text list "Input_注释": 0 '备用'; 1 '备用'; 2 '备用'; 3 '备用'; 4 '备用'; 5 '备用'; 6 '备用'; 7 '备用'; 10 '备用'; 11 '备用'; 12 '备用'; 13 '备用'; 14 '备用'; 15 '备用'; 16 '备用'; 17 '备用'; 20 '紧急停止 / 备用'; 21 '总气压检测 / 备用'; 22 '手动模式 / 备用'; 23 '自动模式 / 备用'; 24 '启动运行按钮 / 备用'; 25 '故障复位按钮 / 备用'; 26 '启动按钮输入 / 备用'; 27 '光幕Ok / RobotReadyToMark'; 30 '旁路钥匙开关'; 31 '备用 / RobotTrayFullToOut'; 32 '变频器Ready / RobotPartInTurner'; 33 '备用 / reserve'; 34 '备用'; 35 '备用'; 36 '备用'; 37 '备用'; 40 '备用'; 41 '备用'; 42 '备用'; 43 '备用'; 44 '备用'; 45 '备用'; 46 '备用'; 47 '备用'; 50 '备用'; 51 '备用'; 52 '备用'; 53 '备用'; 54 '备用'; 55 '备用'; 56 '备用'; 57 '备用'; 200 '10插销缸缩回位磁开 / Communication with Conveyor / 与Conveyor通讯'; 201 '10插销缸伸出位磁开 / Communication with Conveyor / 与Conveyor通讯'; 202 '10测试滑台缸伸出位磁开'; 203 '10测试滑台缸缩回位磁开 / Communication with Conveyor / 与Conveyor通讯'; 204 '10测试升降缸伸出位磁开 / Communication with Conveyor / 与Conveyor通讯'; 205 '10测试升降缸缩回位磁开 / Communication with Conveyor / 与Conveyor通讯'; 206 '10滑台推出缸缩回位磁开 / Communication with Conveyor / 与Conveyor通讯'; 207 '10滑台推出缸伸出位磁开 / Communication with Conveyor / 与Conveyor通讯'; 210 '10下料滑台缸伸出位磁开 / Communication with Conveyor / 与Conveyor通讯'; 211 '10下料滑台缸缩回位磁开 / Communication with Conveyor / 与Conveyor通讯'; 212 '11下料升降缸伸出位磁开 / Communication with Conveyor / 与Conveyor通讯'; 213 '11下料升降缸缩回位磁开 / Communication with Conveyor / 与Conveyor通讯'; 214 '11下料夹爪缸伸出位磁开 / Communication with Conveyor / 与Conveyor通讯'; 215 '11下料夹爪缸缩回位磁开 / Communication with Conveyor / 与Conveyor通讯'; 216 '11废料阻挡缸伸出位磁开 / Communication with Conveyor / 与Conveyor通讯'; 217 '11废料阻挡缸缩回位磁开 / Communication with Conveyor / 与Conveyor通讯'; 222 '10.气密工件到位接近开关信号 / Communication with Conveyor / 与Conveyor通讯'; 223 '10.废料检测信号 / Communication with Conveyor / 与Conveyor通讯'; 224 '11.气密下料工件到位信号 / Communication with Conveyor / 与Conveyor通讯'; 225 '备用 / Communication with Conveyor / 与Conveyor通讯'; 226 '备用 / Communication with Conveyor / 与Conveyor通讯'; 227 '备用 / Communication with Conveyor / 与Conveyor通讯'; 230 '2垂直探针缸伸出位磁开 / Communication with Conveyor / 与Conveyor通讯'; 232 '备用 / Communication with Conveyor / 与Conveyor通讯'; 233 '备用 / Communication with Conveyor / 与Conveyor通讯'; 234 '转盘上料位工件到位信号 / Communication with Conveyor / 与Conveyor通讯'; 235 '备用 / Communication with Conveyor / 与Conveyor通讯'; 236 '备用 / Communication with Conveyor / 与Conveyor通讯'; 240 '2水平探针缸伸出位磁开 / Indexing plate number 3 / 转盘编号3'; 241 '2水平探针缸缩回位磁开 / Indexing plate number 4 / 转盘编号4'; 242 '8升降缸伸出位磁开 / 06.压紧缸原点位磁开'; 243 '8升降缸缩回位磁开 / 06.压紧缸工作位磁开'; 244 '2夹紧缸缩回位磁开 / 06.热烫缸原点位磁开'; 245 '2夹紧缸伸出位磁开 / 06.热烫缸工作位磁开'; 246 '备用 / 02.升降缸原点位磁开'; 247 '备用 / 02.升降缸工作位磁开'; 250 '4齿面凹面转换缸伸出位磁开 / Indexing plate number 1 / 转盘编号1'; 251 '4齿面凹面转换缸缩回位磁开 / Indexing plate number 2 / 转盘编号2'; 252 '4垂直探针缸伸出位磁开 / 上料托盘检测光电1'; 253 '4垂直探针缸缩回位磁开 / 上料皮带挡料1缸工作位磁开'; 254 '4夹紧缸缩回位磁开 / 上料皮带挡料2缸工作位磁开'; 255 '4夹紧缸伸出位磁开 / 上料托盘检测光电2'; 256 '4水平探针缸伸出位磁开 / 02.送料长缸工作位磁开'; 257 '4水平探针缸缩回位磁开 / 02.送料长缸原点位磁开'; 260 '6夹紧缸缩回位磁开 / 02.送料短缸工作位磁开'; 261 '6夹紧缸伸出位磁开 / 01.真空*工作位磁开'; 262 '6水平探针缸伸出位磁开 / 06.热烫缸工作位磁开'; 263 '6水平探针缸缩回位磁开 / 06.热烫缸工作位磁开'; 264 '6垂直探针缸伸出位磁开 / 06.热烫缸工作位磁开'; 265 '6垂直探针缸缩回位磁开 / 06.热烫缸工作位磁开'; 266 '02.转台编码 Bit0 / 06.热烫缸工作位磁开'; 267 '02.转台编码 Bit1 / 06.热烫缸工作位磁开'; 270 '02.转台编码 Bit2 / 06.热烫缸工作位磁开'; 271 '02.转台编码 Bit3 / 06.热烫缸工作位磁开'; 272 '备用 / 06.热烫缸工作位磁开'; 273 '备用 / 06.热烫缸工作位磁开'; 274 '备用 / 06.热烫缸工作位磁开'; 275 '备用 / 06.热烫缸工作位磁开'; 276 '备用 / 06.热烫缸工作位磁开'; 277 '备用 / 06.热烫缸工作位磁开'; 280 '备用 / 06.热烫缸工作位磁开'; 220 '10.气密工件到位光电信号 / Communication with Conveyor / 与Conveyor通讯'; 221 '备用 / Communication with Conveyor / 与Conveyor通讯'; 231 '2垂直探针缸缩回位磁开 / Communication with Conveyor / 与Conveyor通讯'; 237 '转台到位检测接近 / Communication with Conveyor / 与Conveyor通讯'; 281 '备用 / 06.热烫缸工作位磁开'; 282 '备用 / 06.热烫缸工作位磁开'; 283 '备用 / 06.热烫缸工作位磁开'; 284 '备用 / 06.热烫缸工作位磁开'; 285 '备用 / 06.热烫缸工作位磁开'; 286 '07.工件到位信号'; 287 '备用'; 290 '07.插销缸缩回信号'; 291 '07.插销缸伸出信号'; 292 '07.压紧缸缩回信号'; 293 '07.压紧缸伸出信号'; 294 '备用'; 295 '备用'; 296 '07.滑台推进缸伸出信号'; 297 '07.滑台推进缸缩回信号'; 300 '07.下料滑台缸缩回信号'; 301 '07.下料滑台缸伸出信号'; 302 '08.下料升降缸伸出信号'; 303 '08.下料升降缸缩回信号'; 304 '08.下料夹爪缸缩回信号'; 305 '08.下料夹爪缸伸出信号'; 306 '08.下料止挡缸伸出信号'; 307 '08.下料止挡缸缩回信号'; 310 '备用'; 311 '备用'; 312 '备用'; 313 '备用'; 314 '备用'; 315 '备用'; 316 '备用'; 317 '备用'; 74 '备用'; 77 '备用'; 76 '备用'; 75 '备用'; 73 '备用'; 72 '备用'; 71 '备用'; 70 '备用'; 67 '备用'; 66 '备用'; 65 '备用'; 64 '备用'; 63 '备用'; 62 '备用'; 61 '备用'; 60 '备用'; 320 '备用'; 321 '备用'; 322 '备用'; 323 '备用'; 324 '备用'; 325 '备用'; 326 '备用'; 327 '备用'; 330 '备用'; 331 '备用'; 332 '备用'; 333 '备用'; 334 '备用'; 335 '备用'; 336 '备用'; 337 '备用'; 340 '备用'; 341 '备用'; 342 '备用'; 343 '备用'; 344 '备用'; 345 '备用'; 346 '备用'; 347 '备用'; 350 '备用'; 351 '备用'; 352 '备用'; 353 '备用'; 354 '备用'; 355 '备用'; 356 '备用'; 357 '备用'

text list "OutPut_地址": 0 'Q0.0'; 1 'Q0.1'; 2 'Q0.2'; 3 'Q0.3'; 4 'Q0.4'; 5 'Q0.5'; 6 'Q0.6'; 7 'Q0.7'; 10 'Q1.0'; 11 'Q1.1'; 12 'Q1.2'; 13 'Q1.3'; 14 'Q1.4'; 15 'Q1.5'; 16 'Q1.6'; 17 'Q1.7'; 20 'Q2.0'; 21 'Q2.1'; 22 'Q2.2'; 23 'Q2.3'; 24 'Q2.4'; 25 'Q2.5'; 26 'Q2.6'; 27 'Q2.7'; 30 'Q3.0'; 31 'Q3.1'; 32 'Q3.2'; 33 'Q3.3'; 34 'Q3.4'; 35 'Q3.5'; 36 'Q3.6'; 37 'Q3.7'; 40 'Q4.0'; 41 'Q4.1'; 42 'Q4.2'; 43 'Q4.3'; 44 'Q4.4'; 45 'Q4.5'; 46 'Q4.6'; 47 'Q4.7'; 50 'Q5.0'; 51 'Q5.1'; 52 'Q5.2'; 53 'Q5.3'; 54 'Q5.4'; 55 'Q5.5'; 56 'Q5.6'; 57 'Q5.7'; 200 'Q20.0'; 201 'Q20.1'; 202 'Q20.2'; 203 'Q20.3'; 204 'Q20.4'; 205 'Q20.5'; 206 'Q20.6'; 207 'Q20.7'; 210 'Q21.0'; 211 'Q21.1'; 212 'Q21.2'; 213 'Q21.3'; 214 'Q21.4'; 215 'Q21.5'; 216 'Q21.6'; 217 'Q21.7'; 220 'Q22.0'; 221 'Q22.1'; 222 'Q22.2'; 223 'Q22.3'; 224 'Q22.4'; 225 'Q22.5'; 226 'Q22.6'; 227 'Q22.7'; 230 'Q23.0'; 231 'Q23.1'; 232 'Q23.2'; 233 'Q23.3'; 234 'Q23.4'; 235 'Q23.5'; 236 'Q23.6'; 237 'Q23.7'; 240 'Q24.0'; 241 'Q24.1'; 242 'Q24.2'; 243 'Q24.3'; 244 'Q24.4'; 245 'Q24.5'; 246 'Q24.6'; 247 'Q24.7'; 250 'Q25.0'; 251 'Q25.1'; 252 'Q25.2'; 253 'Q25.3'; 254 'Q25.4'; 255 'Q25.5'; 256 'Q25.6'; 257 'Q25.7'; 260 'Q26.0'; 261 'Q26.1'; 262 'Q26.2'; 263 'Q26.3'; 264 'Q26.4'; 265 'Q26.5'; 266 'Q26.6'; 267 'Q26.7'; 270 'Q27.0'; 271 'Q27.1'; 272 'Q27.2'; 273 'Q27.3'; 274 'Q27.4'; 275 'Q27.5'; 276 'Q27.6'; 277 'Q27.7'; 280 'Q28.0'; 281 'Q28.1'; 282 'Q28.2'; 283 'Q28.3'; 284 'Q28.4'; 285 'Q28.5'; 286 'Q28.6'; 287 'Q28.7'; 290 'Q29.0'; 291 'Q29.1'; 292 'Q29.2'; 293 'Q29.3'; 294 'Q29.4'; 295 'Q29.5'; 296 'Q29.6'; 297 'Q29.7'; 67 'Q6.7'; 66 'Q6.6'; 65 'Q6.5'; 64 'Q6.4'; 63 'Q6.3'; 62 'Q6.2'; 61 'Q6.1'; 60 'Q6.0'; 77 'Q7.7'; 76 'Q7.6'; 75 'Q7.5'; 74 'Q7.4'; 73 'Q7.3'; 72 'Q7.2'; 71 'Q7.1'; 70 'Q7.0'; 300 'Q30.0'; 301 'Q30.1'; 302 'Q30.2'; 303 'Q30.3'; 304 'Q30.4'; 305 'Q30.5'; 306 'Q30.6'; 307 'Q30.7'

text list "OutPut_注释": 0 '备用'; 1 '备用'; 2 '备用'; 3 '备用'; 4 '备用'; 5 '备用'; 6 '备用'; 7 '备用'; 10 '备用'; 11 '备用'; 12 '备用'; 13 '备用'; 14 '备用'; 15 '备用'; 16 '备用'; 17 '备用'; 20 '面板.蜂鸣器'; 21 '面板.绿色运行灯'; 22 '面板.故障复位红灯'; 23 '三色塔灯(红)'; 24 '三色塔灯(黄)'; 25 '三色塔灯(绿)'; 26 '启动按钮指示灯'; 27 '日光灯控制'; 30 '总气源开电磁阀'; 31 '旁路中继'; 32 '变频器复位'; 33 '转台电机运行'; 34 '测试探针切换中继'; 35 '备用'; 36 '备用'; 37 '转台到位指示灯'; 40 '抽烟机启动'; 41 '备用'; 42 '备用'; 43 '备用'; 44 '备用'; 45 '备用'; 46 '合格件指示灯'; 47 '疑品件指示灯'; 50 '备用'; 51 '备用'; 52 '备用'; 53 '备用'; 54 '备用'; 55 '备用'; 56 '备用'; 57 '备用'; 200 '2水平探针缸伸出电磁阀'; 201 '2水平探针缸缩回电磁阀'; 202 '2垂直探针缸伸出电磁阀'; 203 '2垂直探针缸缩回电磁阀'; 204 '2夹紧缸伸出电磁阀'; 205 '2夹紧缸缩回电磁阀'; 206 '4齿面凹面转换缸伸出电磁阀'; 207 '4齿面凹面转换缸缩回电磁阀'; 210 '4垂直探针缸伸出电磁阀'; 211 '4垂直探针缸缩回电磁阀'; 212 '4夹紧缸伸出电磁阀'; 213 '4夹紧缸缩回电磁阀'; 214 '4水平探针缸伸出电磁阀'; 215 '4水平探针缸缩回电磁阀'; 216 '6夹紧缸伸出电磁阀'; 217 '6夹紧缸缩回电磁阀'; 220 '6水平探针缸伸出电磁阀'; 221 '6水平探针缸缩回电磁阀'; 222 '6垂直探针缸伸出电磁阀'; 223 '6垂直探针缸缩回电磁阀'; 224 '8升降缸伸出电磁阀'; 225 '8升降缸缩回电磁阀'; 226 '10插销缸伸出电磁阀'; 227 '10插销缸缩回电磁阀'; 230 '10测试滑台缸伸出电磁阀'; 231 '10测试滑台缸缩回电磁阀'; 232 '10测试升降缸伸出电磁阀'; 233 '10测试升降缸缩回电磁阀'; 234 '10滑台推出缸伸出电磁阀'; 235 '10滑台推出缸缩回电磁阀'; 236 '10下料滑台缸伸出电磁阀'; 237 '10下料滑台缸缩回电磁阀'; 240 '11下料升降缸伸出电磁阀'; 241 '11下料升降缸缩回电磁阀'; 242 '11下料夹爪缸伸出电磁阀'; 243 '11下料夹爪缸缩回电磁阀'; 244 '11废料阻挡缸伸出电磁阀'; 245 '11废料阻挡缸缩回电磁阀'; 246 '备用'; 247 '备用'; 250 '备用'; 251 '备用'; 252 '备用'; 253 '备用'; 254 '备用'; 255 '备用'; 256 '备用'; 257 '备用'; 260 '备用'; 261 '备用'; 262 '备用'; 263 '备用'; 264 '备用'; 265 '备用'; 266 '备用'; 267 '备用'; 270 '备用'; 271 '备用'; 272 '备用'; 273 '备用'; 274 '备用'; 275 '备用'; 276 '备用'; 277 '备用'; 280 '备用'; 281 '备用'; 77 '备用'; 76 '备用'; 75 '备用'; 74 '备用'; 73 '备用'; 72 '备用'; 71 '备用'; 70 '备用'; 67 '备用'; 66 '备用'; 65 '备用'; 64 '备用'; 63 '备用'; 62 '备用'; 61 '备用'; 60 '备用'; 304 '备用'; 305 '备用'; 306 '备用'; 307 '备用'

text list "CognexStatusPrompt": 0 'info. ModeOff !'; 1 'info. Online'; 2 'info. Programming'; 3 'info. Discrete Offline'; 4 'info. Comm. Offline'; 5 'info. triger cycle Wait for Triger Ack signal'; 6 'info. triger cyclle Wait for inspection completed signal'; 7 'info. wait for triger ready signal!'; 8 'info. Wait for offline to load job!'; 9 'info. Wait for job load completed!'; 10 'info. Triger result Pass !'; 11 'info. JobLoad OK !'; 12 'info.6'; 13 'info.5'; 14 'info.4'; 15 'info.3'; 16 'info.1'; 17 ''; 18 ''; 19 ''; 20 ''; 21 'xx'; 22 ''; 23 ''; 24 ''; 25 ''; 26 ''; 27 ''; 28 ''; 29 ''; 30 ''; 31 'info.'; 32 'Err. Connnect Err, Pls Reset!'; 33 'Err. Job load fail!'; 34 'Err. Triger Result Fail !'; 35 ''; 36 ''; 37 ''; 38 ''; 39 ''; 40 ''; 41 ''; 42 ''; 43 'info.7'; 44 'info.6'; 45 'info.5'; 46 'info.4'; 47 'info.3'; 48 'info.1'; 49 ''; 50 ''; 51 'xx'; 52 ''; 53 ''; 54 ''; 55 ''; 56 ''; 57 ''; 58 ''; 59 ''; 60 ''; 61 ''; 62 ''; 63 'Err.'; 30000 'no info.'

text list "MotionCtrl_PLCOpen_Status": 0 'EMMode'; 1 'ServoProhibited'; 2 'RestartRequired'; 3 'ServoLostRef'; 4 'NotActivated'; 5 'Position...'; 6 'Homeing...'; 7 'Jog...'; 8 'ServoReady'; 9 'Mode off!'; 10 ''; 11 ''; 12 ''; 13 ''; 14 ''; 15 ''; 16 ''; 17 ''; 18 ''; 19 ''; 20 ''; 21 ''; 22 ''; 23 ''; 24 ''; 25 ''; 26 ''; 27 ''; 28 ''; 29 ''; 30 ''; 31 'Info'; 32 'NotEnable'; 33 'NotActivated'; 34 'Servo controller alarm present'; 35 'Servo Controller InPosition Signal Err'; 36 'Internal_Err'; 37 'Configuration error'; 38 'Servo controller not ready!'; 39 'Low SW limit reached'; 40 'Low SW limit exceeded'; 41 'High SW limit reached'; 42 'High SW limit exceeded'; 43 'Low HW limit switch has been approached'; 44 'High HW limit switch has been approached'; 45 ''; 46 ''; 47 ''; 48 ''; 49 ''; 50 ''; 51 ''; 52 ''; 53 ''; 54 ''; 55 ''; 56 ''; 57 'info.6'; 58 'info.7'; 59 'info.1'; 60 'info.2'; 61 'info.3'; 62 'info.4'; 63 'info.5'; 3000 'no info.'; 2999 'S7 Connect Fail !'

text list "SC_Prompt_Status": 0 'info. Mode = Off !'; 1 'info. Serial Communication started!'; 2 'info. Send Starting ...'; 3 'info. Send OK, Wait for Response'; 4 'info. Recv OK ...'; 5 'info. Wait for Command Off'; 6 'info. time out retrying !'; 7 ''; 8 ''; 9 ''; 10 'info.'; 11 ''; 12 ''; 13 ''; 14 ''; 15 'xx'; 16 'info.1'; 17 'info.3'; 18 'info.4'; 19 'info.5'; 20 'info.6'; 21 ''; 22 ''; 23 ''; 24 ''; 25 ''; 26 ''; 27 ''; 28 ''; 29 ''; 30 ''; 31 'info'; 32 'Err. Send FB Error !'; 33 'Err. Recv FB Error !'; 34 'Err. ResponseTimeOut, Retrying !'; 35 'Err. NotReady!'; 36 'Err. Communication time out ! 10s'; 37 ''; 38 ''; 39 ''; 40 ''; 41 ''; 42 ''; 43 'Err.'; 44 ''; 45 ''; 46 ''; 47 ''; 48 ''; 49 ''; 50 'info.5'; 51 'info.6'; 52 'info.7'; 53 ''; 54 ''; 55 ''; 56 ''; 57 ''; 58 'info.1'; 59 'info.3'; 60 'info.4'; 61 ''; 62 ''; 63 'xx'; 30000 'no info.'

text list "Print": 0 'info. ModeOff !'; 1 'info. Online'; 2 'info. Programming'; 3 'info. Discrete Offline'; 4 'info. Comm. Offline'; 5 'info. triger cycle Wait for Triger Ack signal'; 6 'info. triger cyclle Wait for inspection completed signal'; 7 'info. wait for triger ready signal!'; 8 'info. Wait for offline to load job!'; 9 'info. Wait for job load completed!'; 10 'info. Triger result Pass !'; 11 'info. JobLoad OK !'; 12 'info.6'; 13 'info.5'; 14 'info.4'; 15 'info.3'; 16 'info.1'; 17 ''; 18 ''; 19 ''; 20 ''; 21 'xx'; 22 ''; 23 ''; 24 ''; 25 ''; 26 ''; 27 ''; 28 ''; 29 ''; 30 ''; 31 'info.'; 32 'Err. Connnect Err, Pls Reset!'; 33 'Err. Job load fail!'; 34 'Err. Triger Result Fail !'; 35 'Err.Character String Change Error'; 36 'Err.Print Error'; 37 'Err.Program Change Error'; 38 'Err.Character String Read Error'; 39 ''; 40 ''; 41 ''; 42 ''; 43 'info.7'; 44 'info.6'; 45 'info.5'; 46 'info.4'; 47 'info.3'; 48 'info.1'; 49 ''; 50 ''; 51 'xx'; 52 ''; 53 ''; 54 ''; 55 ''; 56 ''; 57 ''; 58 ''; 59 ''; 60 ''; 61 ''; 62 ''; 63 'Err.'; 30000 'no info.'

text list "KeyenceMD_X_StatusPrompt": 0 'info. ModeOff !'; 1 'info.Triger not ready!'; 2 'info. Shutter Closed!'; 3 'info. Profinet communication not started'; 4 'info. Clearing Error'; 5 'info. Main Step is running, Busy'; 6 'info. wait user command off!'; 7 'info. JobLoad OK !'; 8 'info. Printing !'; 9 'info. Prog Loading!'; 10 'info. Requesting parameter'; 11 'info. Ok To Start'; 12 ''; 13 ''; 14 ''; 15 ''; 16 ''; 17 ''; 18 ''; 19 ''; 20 ''; 21 ''; 22 ''; 23 ''; 24 ''; 25 ''; 26 ''; 27 ''; 28 ''; 29 ''; 30 ''; 31 'info.'; 32 'Err. Connnect Err, Pls Reset!'; 33 'Err. Job load fail!'; 34 'Err.Character String Change Error'; 35 'Err.Print Error'; 36 'Err.Program Change Error'; 37 'Err.Character String Read Error'; 38 ''; 39 ''; 40 ''; 41 ''; 42 'info.7'; 43 'info.6'; 44 'info.5'; 45 'info.4'; 46 'info.3'; 47 'info.1'; 48 ''; 49 ''; 50 'xx'; 51 ''; 52 ''; 53 ''; 54 ''; 55 ''; 56 ''; 57 ''; 58 ''; 59 ''; 60 ''; 61 ''; 62 ''; 63 'Err.'

text list "模式": 0 '单机'; 1 '联机'

text list "打标": 0 '打标'; 1 '不打标'

text list "Siemens_V90_FaultCodeText": 0 '正常'; 1000 '内部软件错误'; 1001 '浮点例外'; 1002 '内部软件错误'; 1003 '访问存储器时出现应答延迟'; 1010 '驱动类型不明'; 1011 '(N)下载中断'; 1012 '(N)项目转化出错'; 1015 '内部软件错误'; 1023 '内部软件超时'; 1030 '控制权下的生命符号出错'; 1031 '“远程模式关”下的生命符号出错'; 1033 '单位转换：参考参数无效'; 1034 '单位转换：参考值更改后参数值计算失败'; 1036 'ACX：缺少参数备份文件'; 1038 'ACX：载入参数备份文件失败'; 1039 'ACX：写入参数备份文件失败'; 1040 '需要备份参数并重新上电'; 1041 '需要备份参数'; 1042 '下载项目时的参数出错'; 1043 '在项目下载时出现严重错误'; 1044 'CU：描述数据出错'; 1050 '存储卡和设备不兼容'; 1054 'CU:超出系统极限'; 1055 'CU：内部错误（应用和端口的SYNO不相同）'; 1056 'CU：内部错误（参数组时钟周期已经分配，但有偏差）'; 1058 'CU：内部错误（拓扑结构中没有从站）'; 1059 'CU：内部错误（端口不存在）'; 1060 'CU：内部错误（参数组不存在）'; 1061 'CU：内部错误（应用未知）'; 1063 'CU：内部错误（PDM）'; 1068 'CU：数据存储器溢出'; 1070 '正在向存储卡进行项目/固件下载'; 1072 '从备份文件中修复存储卡'; 1105 'CU：存储器容量不足'; 1106 'CU：存储器容量不足'; 1107 'CU：保存到非易失性存储器的操作失败'; 1110 'CU：一个控制单元上不止一个SINAMICSG'; 1111 'CU：不允许驱动设备混合运行'; 1112 'CU:功率单元非法'; 1120 '初始化端口失败'; 1122 '测量探头输入端的频率过高'; 1123 '功率单元不支持数字输入/输出端'; 1150 'CU：超过了某一驱动对象类型的实例数'; 1151 'CU：超出了某一类别驱动对象的数量'; 1200 'CU:时间片管理内部软件错误'; 1205 'CU：时间片溢出'; 1221 'CU：基本周期太小'; 1222 'CU：基本时钟周期太小（没有用于通讯的计算时间）'; 1223 'CU：采样时间不一致'; 1250 'CU：CU-EEPROM只读数据出错'; 1255 'CU:插件板EEPROM只读数据出错'; 1325 '拓扑结构：设定拓扑结构中不包含该组件号'; 1340 '拓扑结构：一个支路上的组件过多'; 1354 '拓扑结构：实际拓扑结构存在错误的组件'; 1355 '拓扑结构：实际拓扑结构已更改'; 1360 '拓扑结构：实际拓扑结构非法'; 1375 '组件：两个组件之间实际拓扑结构连接重复'; 1380 '拓扑结构：实际拓扑结构损坏的EEPROM'; 1451 '设定拓扑结构无效'; 1470 '拓扑结构：发现设定拓扑结构环形连接'; 1475 '拓扑结构：两个组件之间设定拓扑结构连接重复'; 1506 'BICO:无标准报文'; 1510 'BICO：信号源不是浮点'; 1511 'BICO：连接有不同定标'; 1512 'BICO：没有定标'; 1513 'BICO：不同驱动对象之间的连接有不同定标'; 1514 '(F)BICO：在重新连接期间写入时出错'; 1515 'BICO:不允许写入参数，因为控制权有效'; 1600 'SICU：STOPA被触发'; 1611 'SICU：某一监控通道故障'; 1612 'SICU:并联功率单元上STO输入不同'; 1625 'SICU：安全数据中生命符号出错'; 1630 'SICU:制动控制出错'; 1649 'SICU:内部软件错误'; 1650 'SICU:必须进行验收测试'; 1651 'SICU：安全时间片同步失败'; 1652 'SICU:非法的监控周期'; 1653 'SICU:PROFIBUS/PROFINET配置出错'; 1655 'SICU：监控功能的对比'; 1656 'SICU：电机模块参数出错'; 1657 'SICU:PROFIsafe报文号无效'; 1658 'SICU:PROFIsafe报文号不一致'; 1659 'SICU：参数的写入任务被绝'; 1660 'SICU：不支持安全功能'; 1661 'SICU:安全输入端模拟激活'; 1663 'SICU：SI参数复制被拒绝'; 1664 'SICU：无自动固件升级'; 1665 'SICU:系统故障'; 1670 'SI运动：编码器模块参数设置无效'; 1671 'SI运动：编码器参数设置出错'; 1672 'SICU：电机模块软件/硬件不兼容'; 1673 'SI运动：编码器模块软件/硬件不兼容'; 1674 'SI运动CU：PROFIsafe报文不支持安全功能'; 1680 'SI运动CU：安全监控校验和错误'; 1681 'SI运动CU：参数值误'; 1682 'SI运动CU：不支持监控功能'; 1683 'SI运动CU：缺少SOS/SLS使能'; 1684 'SI运动：Safely-LimitedPosition极限值混淆'; 1685 'SI运动CU：Safely-LimitedSpeed的极限值过大'; 1686 'SI运动：凸轮位置参数设置出错'; 1687 'SI运动：SCA(SN)模数值设定出错'; 1688 'SI运动CU：不允许实际值同步'; 1690 'SI运动:NVRAM上的数据备份问题'; 1692 'SI运动CU：无编码器时参数值错误'; 1694 'SI运动CU:电机模块的固件版本低于控制单元'; 1695 '5(F)SI运动：编码器模块被更换'; 1786 'SCC信号被修改'; 1787 'SBT电机类型不同'; 1910 '现场总线设定值超时'; 1911 'PB/PN等时同步周期故障'; 1912 'PB/PN等时同步中生命符号出错'; 1913 'COMMINT：生命符号监控时间结束'; 1914 'COMMINT：配置监控时间结束'; 1915 'PB/PN同步运行，驱动对象1生命符号出错'; 1950 'PB/PN等时同步失败'; 2080 '跟踪：参数设置由于单位转换被删除'; 2151 'OA:内部软件错误'; 2152 'OA:存储器容量不够'; 3000 '操作时的NVRAM错误'; 3001 'NVRAM校验和出错'; 3500 'TM：初始化'; 3505 '模拟输入端断线'; 5055 '并联电路：功率单元代码号非法'; 5056 '并联电路：功率单元EPROM版本不同'; 5057 '并联电路：功率单元固件版本不同'; 5058 '并联电路：VSMEEPROM版本不同'; 5059 '并联电路：VSM固件版本不同'; 5060 '并联电路：功率单元固件版本不兼容'; 5061 '整流单元VSM数量'; 5064 '并联：脉冲同步错误'; 5118 '超出预充电接触器同步监控时间'; 5119 '超出分路接触器同步监控时间'; 6000 '整流单元：预充电监控时间已结束'; 6010 '整流单元：运行中缺少功率单元EP24V'; 6050 '整流单元：不支持非调节模式'; 6052 '整流单元：不支持滤波器温度检测'; 6100 '整流单元：由于主电源欠电压断路'; 6200 '整流单元：一个或者多个主电源相位故障'; 6210 '整流单元：总电流过高'; 6211 '整流单元：总电流过高'; 6261 '整流单元：输入滤波器温度持续过高'; 6262 '整流单元：接通时输入滤波器内的温度开关打开'; 6300 '整流单元：在接通时输入电压过高'; 6310 '输入电压(p0210)参数设定错误'; 6311 '整流单元：输入电压（p0210）故障'; 6320 '主站/从站：4通道多路转换器控制无效'; 6321 '主站/从站：6通道多路换器控制无效'; 6504 '整流单元：孤岛电网同步失败'; 6700 '整流单元：负载时接通电源接触器'; 6850 '整流单元：短路时间过长'; 6851 '整流单元：分布式整流单元的电源监控已触发'; 6855 '整流单元：输入滤波器监控已响应'; 6906 '制动模块内部故障信息'; 6907 '制动模块内部过热'; 6908 '制动模块内部过热/断路'; 6909 '制动模块内部Uce故障'; 6922 '制动电阻断相'; 7011 '驱动：电机超温'; 7013 '驱动：电机温度模型配置故障'; 7016 '驱动：电机温度传感器的故障信息'; 7018 '超出附加温度故障阈值'; 7080 '驱动：闭环控制参数出错'; 7082 '宏文件：无法执行'; 7083 '宏文件：找不到ACX文件'; 7084 '宏文件：未满足WaitUntil的条件'; 7085 '驱动：开环控制/闭环控制参数被更改'; 7086 '单位转换:由于参考值改变而超出参数极限'; 7087 '驱动：在设定的脉冲频率下无法进行无编码器运行'; 7088 '单位转换:由于单位转换而超出参数极限'; 7090 '驱动：转矩上限小于下限'; 7100 '驱动：采样时间不可复位'; 7110 '驱动：采样时间和基本周期不匹配'; 7220 '驱动：缺少“通过PLC控制”'; 7300 '驱动：缺少电源接触器反馈信息'; 7311 '电机旁路开关'; 7312 '电源旁路开关'; 7320 '驱动：自动重启中断'; 7331 '捕捉再启动:不支持该功能'; 7403 '驱动：达到直流母线电压阈值下限'; 7404 '驱动：达到直流母线电压阈值上限'; 7405 '驱动：低于动能缓冲下的最低转速'; 7406 '驱动：超出动能缓冲状态下最大持续时间'; 7407 '驱动：不允许Vdc降低'; 7410 '驱动：电流环输出受限'; 7411 '驱动：磁通控制器输出受限'; 7412 '驱动：换向角出错（电机模型）'; 7413 '驱动：换向角出错（磁极位置检测）'; 7414 '驱动：编码器序列号改变'; 7417 '驱动脉冲方式不合理（电机模型）'; 7419 '驱动：电流设定值滤波器自适应配置不一致'; 7420 '驱动：电流设定值滤波器固有频率>香农频率'; 7421 '驱动：转速滤波器固有频率>香农频率'; 7422 '驱动：参考模型固有频率>香农频率'; 7423 '驱动：APC滤波器固有频率>香农频率'; 7425 '驱动：APC转速极限监控时间超期'; 7426 '工艺控制器实际值达到极限值'; 7429 '驱动：无编码器时不支持DSC'; 7430 '驱动：无法切换到转矩开环运行'; 7431 '驱动：无法切换到无编码器运行'; 7432 '驱动：电机无过压保护'; 7433 '驱动：无法切换到带编码器运行，因为编码器没有解除驻留'; 7434 '驱动：无法在脉冲使能时改变旋转方向'; 7435 '(N)驱动：无编码器的矢量控制，斜坡函数发生器设置错误'; 7439 '驱动:不支持该功能'; 7442 '位置环：多圈分辨率和模数范围不匹配'; 7443 '位置环：参考点坐标超出允许范围'; 7446 '负载变速箱：无法复位位置跟踪'; 7447 '负载变速箱：位置跟踪超出最大实际值'; 7448 '负载变速箱：位置跟踪线性轴超出最大范围'; 7449 '负载变速箱：位置跟踪当前位置在公差范围之外'; 7450 '位置环:静态监控已响应'; 7451 '位置环:定位监控已响应'; 7452 '位置环:跟随误差过大'; 7453 '位置环：位置实际值处理出错'; 7458 'EPOS：未找到参考点凸轮'; 7459 'EPOS：不存在零脉冲'; 7460 'EPOS：未找到参考点凸轮结束点'; 7475 'EPOS：目标位置<运行范围起始处'; 7476 'EPOS：目标位置>运行范围结束处'; 7481 'EPOS：轴位置<负软件限位开关'; 7482 'EPOS：轴位置>正软件限位开关'; 7484 'EPOS：固定挡块在监控窗口之外'; 7485 'EPOS：未到达固定挡块'; 7488 'EPOS：无法相对定位'; 7490 '(N)EPOS：运行时取消使能'; 7491 'EPOS：到达负停止凸轮'; 7492 'EPOS：到达正停止凸轮'; 7493 '位置环：位置实际值的值范围溢出'; 7494 '位置环：在运行时切换驱动数据组'; 7499 'EPOS：沿错误方向到达反向凸轮'; 7500 '驱动：未定义功率单元数据组PDS'; 7501 '驱动：未定义电机数据组MDS'; 7502 '驱动：未定义编码器数据组EDS'; 7503 'EPOS：沿错误运行方向逼近停止凸轮'; 7510 '驱动：驱动数据组中有相同的编码器'; 7511 '驱动：编码器多次使用'; 7512 '驱动：无法设定编码器数据组转换参数'; 7515 '驱动：功率单元和电机连接错误'; 7516 '驱动：重新调试数据组'; 7517 '驱动：编码器数据组转换参数设置错误'; 7518 '驱动：电机数据组转换参数设置错误'; 7551 '驱动编码器：没有换向角信息'; 7552 '驱动编码器：不支持编码器配置'; 7553 '驱动编码器：不支持编码器模块配置'; 7555 '驱动编码器：位置跟踪配置'; 7556 '测量变速箱：位置跟踪超出最大实际值'; 7560 '驱动编码器：线数不是二的幂次方'; 7561 '驱动编码器：多圈线数不是二的幂次方'; 7562 '驱动编码器：增量编码器无法进行位置跟踪'; 7563 '驱动编码器：XIST1_ERW配置错误'; 7575 '驱动：电机编码器未就绪'; 7599 '编码器1：无法校准'; 7600 '编码器2：无法校准'; 7601 '编码器3：无法校准'; 7800 '驱动：没有功率单元'; 7801 '驱动：电机过电流'; 7802 '驱动：整流单元或者功率单元未就绪'; 7805 '(N)整流单元：功率单元过载I2t'; 7807 '驱动：检测出短路/接地'; 7808 'HF阻尼器：阻尼未就绪'; 7810 '驱动：功率单元EEPROM无额定数据'; 7815 '驱动：功率单元已修改'; 7826 '驱动：模拟运行的直流母线电压过高'; 7840 '驱动：缺少整流单元运行'; 7841 '驱动：取消整流单元运行'; 7860 '外部故障1'; 7861 '外部故障2'; 7862 '外部故障3'; 7890 '内部电压保护/内部电枢短路和STO生效'; 7900 '驱动：电机堵转/转速环到达挡块'; 7901 '驱动：电机转速过快'; 7902 '驱动：电机失步'; 7907 '内部电枢短路：在删除脉冲以后，电机端子电位不再隔离'; 7908 '内部电枢短路生效'; 7909 '内部电压保护：只有上电后才失效'; 7913 '励磁电流超出公差'; 7914 '磁通超出公差'; 7923 '驱动：转矩/转速过小'; 7924 '驱动：转矩/转速过大'; 7925 '驱动：转矩/转速超出公差'; 7928 '内部电压保护触发'; 7930 '驱动：制动控制出错'; 7934 '(N)驱动：S120Combi电机抱闸的配置'; 7935 '(N)驱动：电机抱闸配置错误'; 7937 '(N)驱动：电机模型与外部转速的转速偏差'; 7940 '“主电源-驱动”同步：同步故障'; 7950 '驱动：电机参数出错'; 7955 '驱动：电机已经更改'; 7956 '驱动：电机代码与电机列表不匹配'; 7963 '驱动：摩擦特性曲线记录取消'; 7966 '驱动：检查换向角'; 7967 '驱动：编码器自动调校出错'; 7968 '驱动：Lq-Ld测量出错'; 7969 '驱动：磁极位置检测出错'; 7970 '驱动：编码器自动调校出错'; 7982 '驱动：旋转检测编码器测试'; 7983 '驱动：旋转检测饱和特性曲线'; 7984 '驱动：转速环优化，转动惯量异常'; 7985 '驱动：转速环优化（振荡测试）'; 7986 '驱动：旋转检测，斜坡函数发生器异常'; 7988 '驱动：旋转检测未选择配置'; 7989 '驱动：旋转检测，漏电感（q方向）异常'; 7990 '驱动：电机数据检测出错'; 7993 '驱动：旋转磁场方向或者编码器实际值反向出错'; 7994 '(F,N)驱动：未执行电机数据检测'; 7995 '驱动：磁极位置检测失败'; 7996 '驱动：未进行磁极位置检测'; 8000 'TB：电源+/-15V出错'; 8010 'TB：模拟数字转换器'; 8500 'COMMBOARD：配置监控时间结束'; 8501 'COMMBOARD:设定值超时'; 8502 'COMMBOARD：生命符号监控时间结束'; 8510 'COMMBOARD：发送配置数据无效'; 8701 'CAN：NMT状态切换'; 8702 'CAN:RPDO超时'; 8703 'CAN：超过了驱动对象最大数量'; 8751 '(N)CAN：报文丢失'; 13009 'OA应用程序许可未授权'; 13010 '功能模块许可未授权'; 13020 '控制系统中的授权不够'; 13100 '专有技术保护：复制保护故障'; 13101 '专有技术保护：复制保护无法激活'; 13102 '专有技术保护：受保护数据的一致性错误'; 30001 '功率单元：过电流'; 30002 '功率单元：直流母线过电压'; 30003 '功率单元：直流母线欠压'; 30004 '功率单元：逆变器散热器过热'; 30005 '功率单元：I2t过载'; 30006 '功率单元：可控硅控制板'; 30008 '功率单元：循环数据生命符号出错'; 30012 '功率单元：散热器温度传感器断线'; 30013 '功率单元：散热器温度传感器短路'; 30015 '功率单元：电机馈电电缆断相'; 30016 '(N)功率单元：负载电源关闭'; 30017 '功率单元：硬件电流限制响应过于频繁'; 30020 '功率单元：不支持该组态'; 30021 '功率单元：接地'; 30022 '功率单元：U_ce监控'; 30024 '功率单元：热模型过热'; 30025 '功率单元：芯片过热'; 30027 '功率单元：直流母线预充电时间监控'; 30030 '功率单元：内部空间过热报警'; 30035 '功率单元：进风过热'; 30036 '功率单元：内部空间过热'; 30037 '功率单元：整流器过热'; 30039 '功率单元：电容器风扇故障'; 30040 '功率单元：24/48V欠电压'; 30043 '功率单元：24/48V过压'; 30045 '功率单元：电源欠电压'; 30047 '冷却单元：冷却剂体积流量太低'; 30048 '功率单元：外部风扇损坏'; 30050 '功率单元：24V电源过电压'; 30052 'EEPROM数据错误'; 30053 'FPGA数据错误'; 30059 '功率单元：内部风扇损坏'; 30060 '预充电接触器状态监控'; 30061 '旁路接触器状态监控'; 30070 '功率单元不支持所要求的周期'; 30071 '功率单元没有接收到新的实际值'; 30072 '不可再向功率单元传送设定值'; 30074 '控制单元和功率模块之间的通讯出现故障'; 30080 '功率单元：电流提升过快'; 30081 '功率单元：开关操作过于频繁'; 30105 '功率单元：实际值采集出错'; 30314 '功率单：24V电源因PM过载'; 30600 'SIMM:STOPA被触发'; 30611 'SIMM:某一监控通道故障'; 30625 'SIMM：在安全数据中生命符号出错'; 30630 'SIMM:制动控制出错'; 30631 '制动控制：外部打开有效'; 30649 'SIMM:内部软件错误'; 30650 'SIMM:必须进行验收测试'; 30651 'SIMM：与控制单元的同步失败'; 30652 'SIMM:监控周期时间错误'; 30655 'SIMM：监控功能的对比'; 30656 'SIMM：电机模块参数出错'; 30657 'SICU:PROFIsafe报文号无效'; 30659 'SIMM：参数的写入任务被拒绝'; 30662 '内部通讯故障'; 30664 '启动阶段出现故障'; 30665 'SIMM:系统故障'; 30674 'SI运动MM：PROFIsafe报文不支持安全功能'; 30680 'SIMotionMM：安全监控校验和错误'; 30681 'SI运动MM：参数值错误'; 30682 'SI动MM：不支持监控功能'; 30683 'SI运动MM：缺少SOS/SLS使能'; 30684 'SI运动MM：Safely-LimitedPosition极限值混淆'; 30685 'SI运动MM：Safely-LimitedSpeed极限值过大'; 30688 'SI运动MM：实际值同步出错'; 30692 'SI运动MM：无编码器时参数值错误'; 30802 '功率单元：时间片溢出'; 30804 '功率单元：CRC'; 30805 '功率单元：EPROM校验和不正确'; 30809 '功率单元：开关信息无效'; 30850 '功率单元：内部软件错误'; 30899 '功率单元：不明故障'; 30903 '功率单元：出现I2C总线故障'; 30907 '功率单元：FPGA配置失败'; 30950 '功率单元：内部软件错误'; 34207 'VSM：超出温度故障阈值'; 34802 'VSM：时间片溢出'; 34803 'VSM：存储器测试'; 34804 'VSM：CRC'; 34805 'VSM：EPROM校验和不正确'; 34806 'VSM:初始化'; 34850 'VSM：内部软件错误'; 34899 'VSM：不明故障'; 34950 'VSM：内部软件错误'; 35000 'TM54F:采样时间无效'; 35001 'TM54F:参数值无效'; 35002 'TM54F:调试模式被拒'; 35003 'TM54F:需要在控制单元上进行应答'; 35011 'TM54F：驱动对象编号分配错误'; 35013 'TM54F：强制故障检查出错'; 35040 'TM54F：24V欠电压'; 35043 'TM54F：24V过电压'; 35051 'TM54F:某一监控通道故障'; 35052 'TM54F：内部硬件故障'; 35053 'TM54F:超出温度故障阈值'; 35151 'TM54F:差异故障'; 35152 'TM54F：内部软件错误'; 35220 'TM：达到信号输出的极限频率'; 35221 'TM：“设定-实际”差值超出公差'; 35222 '(F,N)TM：编码器线数错误'; 35230 'TM：硬件故障'; 35804 'TM:CRC'; 35899 'TM：不明故障'; 35950 'TM：内部软件错误'; 36207 '集线器：组件过热故障'; 36214 '集线器：24V电源过电压故障'; 36216 '集线器：24V电源欠电压故障'; 36804 '集线器：校验和错误'; 36899 '集线器：不明故障'; 36950 '集线器：内部软件错误'; 37001 'HF阻尼器：过电流'; 37002 'HF阻尼器：阻尼电压过高'; 37003 'HF阻尼器：没有建立阻尼电压'; 37004 'HF阻尼器：散热器过热'; 37005 'HF阻尼器：过载I2t'; 37012 'HF阻尼器：散热器的温度探头断线'; 37013 'HF阻尼器：散热器的温度探头短路'; 37024 'HF阻尼器：热模型超温'; 37025 'HF阻尼器：芯片过热'; 37036 'HF阻尼器：内部空间超温'; 37040 'HF阻尼器：24V欠电压'; 37043 'HF阻尼器：24V过电压'; 37045 'HF阻尼器：电源欠电压'; 37050 'HF阻尼器：24V过电压故障'; 37052 'HF阻尼器：EEPROM数据错误'; 37311 'HF电抗器：散热器超温'; 37313 'HF电抗器：超温或风扇故障'; 37804 'HF阻尼器：CRC'; 37805 'HF阻尼器：EPROM校验和不正确'; 37820 'HF阻尼器：报文错误'; 37835 'HF阻尼器：循环数据传送失败'; 37837 'HF阻尼器：组件故障'; 37845 'HF阻尼器：循环数据传送失败'; 37850 'HF阻尼器：内部软件错误'; 37851 'HF阻尼器(CU)：缺少生命符号'; 37860 'HF阻尼器(CU)：报文错误'; 37875 'HF阻尼器(CU)：电源电压故障'; 37885 'HF阻尼器(CU)：循环数据传送失败'; 37887 'HF阻尼器(CU)：组件故障'; 37895 'HF阻尼器(CU)：交互循环数据传送失败'; 37896 'HF阻尼器(CU)：组件属性不一致'; 37899 'HF阻尼器：不明故障'; 37903 'HF阻尼器：出现I2C总线故障'; 37950 'HF阻尼器：内部软件错误'; 40799 'CX32：超出了定义的传输结束点'; 49150 '冷却单元：出现故障'; 49151 '冷却单元：导热性超出故障阈值'; 49152 '冷却单元：缺少接通指令反馈信息'; 49153 '3冷却单元：冷却液流量过低'; 49154 '冷却单元：出现泄露'; 49155 '冷却单元：功率栈适配器固件版本太旧'; 49156 '冷却单元：冷却液温度超出故障阈值'; 49170 '冷却单元：出报警'

text list "Siemens_V90_ServoStatus": 0 'A00. Controller Stopped'; 1 'A01. Controller Halt'; 2 'A02. Wait for targetPos Reached!'; 3 'A03. Wait for target pos in Band!'; 4 'A04. ModeOff !'; 5 'A05. Permit = off'; 6 'A06. Ready to start'; 7 'A07. Alarm Present'; 8 'A10. Wait for StandStil (check p1226 )'; 9 'A11. forbid axis to forward !'; 10 'A12. forbid axis to backward !'; 11 'A13. Home Seek Started'; 12 'A14. Start Work home process'; 13 'A15. Start Position process!'; 14 'A16. StartTraversingBlock'; 15 'A17. Start Jog movement'; 16 'A20. Start Torque Control Mode'; 17 'A21. Executing parameter communication..'; 18 'A22. TrackIngModeActive'; 19 'A23. Ref = ON, Leaving away Ref Pos !'; 20 'A24.'; 21 'A25.'; 22 'A26.'; 23 'A27.'; 24 'A30.'; 25 'A31'; 26 'A32'; 27 'A33'; 28 'A34'; 29 'A35'; 30 'A36'; 31 'A37'; 32 'E00. Connnect Err, Pls Reset!'; 33 'E01. DriveDisabled by user'; 34 'E02. PLC is sending init para to Drive!'; 35 'E03. Control via PLC Error, Pls check V-Assistant'; 36 'E04. Drive Not Ready For Switch ON, Check DC Supply'; 37 'E05. Drive Enable Failue'; 38 'E06. Fault Present !'; 39 'E07. Reference sensor fault, pls check !'; 40 'E10. Record Communication Error'; 41 'E11. End of Motion fault present'; 42 'E12. Cmd end of time Out !'; 43 'E13. Controller X8.DI3.CWL = Off, pls Check !'; 44 'E14. Controller X8.DI2.CCWL = Off, pls Check!'; 45 'E15.CTRL_IN.RefSource not set !'; 46 'E16. X8.DI4.EMOK = Off,pls Check !'; 47 'E17. SetValuePosition too small !'; 48 'E20. SetValuePosition too large !'; 49 'E21. SetValueVelocity too large !'; 50 'E22'; 51 'E23'; 52 'E24'; 53 'E25'; 54 'E26'; 55 'E27'; 56 'E30'; 57 'E31'; 58 'E32'; 59 'E33'; 60 'E34'; 61 'E35'; 62 'E36'; 63 'E37'

text list "RoundTableV2Prompt_Status": 0 'A00. Not OkToRotate, Pls Reset!'; 1 'A01.'; 2 'A02.'; 3 'A03.'; 4 'A04. ModeOff !'; 5 'A05.'; 6 'A06. Ready to start'; 7 'A07.'; 8 'A10.'; 9 'A11.'; 10 'A12.'; 11 'A13.'; 12 'A14.'; 13 'A15.'; 14 'A16.'; 15 'A17.'; 16 'A20.'; 17 'A21.'; 18 'A22.'; 19 'A23.'; 20 'A24.'; 21 'A25.'; 22 'A26.'; 23 'A27.'; 24 'A30.'; 25 'A31'; 26 'A32'; 27 'A33'; 28 'A34'; 29 'A35'; 30 'A36'; 31 'A37'; 32 'E00. Running time Out( 2s)'; 33 'E01. Inverter is not ready !'; 34 'E02. Two arrival sensor both are On , Pls check !'; 35 'E03. Not OkToRotate !'; 36 'E04'; 37 'E05'; 38 'E06'; 39 'E07'; 40 'E10'; 41 'E11'; 42 'E12'; 43 'E13'; 44 'E14'; 45 'E15'; 46 'E16'; 47 'E17'; 48 'E20'; 49 'E21'; 50 'E22'; 51 'E23'; 52 'E24'; 53 'E25'; 54 'E26'; 55 'E27'; 56 'E30'; 57 'E31'; 58 'E32'; 59 'E33'; 60 'E34'; 61 'E35'; 62 'E36'; 63 'E37'; 30000 'no info.'

text list "机器人动作号": 1 '动作1'; 2 '动作2'; 3 '动作3'; 4 '动作4'; 5 '动作5'

text list "层号": 1 '第1层'; 2 '第2层'; 5 '选择层数'

text list "DB_PromptFree": 0 '气缸操作被禁止，请检查安全条件！'; 1 '设备处于单步模式，请注意安全！'; 2 '设备已经开始清空，请等待！'; 3 '等待循环结束，暂停自动模式中！'; 4 '开始安全门旁路,等待各流程结束!'; 5 '请启动设备！'; 6 '模式来自触摸屏，调试中！'; 7 '光幕被遮,注意安全!'; 8 '请摁下自动模式启动按钮！'; 9 '请求上位机参数录入...'; 10 '请开始换夹具...'; 11 '请求上位机参数录入...'; 12 '换爪运行中'; 13 '水平方向钻入运行中'; 14 '向上方向钻入运行中'; 15 '向下方向钻入运行中'; 16 '检查钻头运行中'; 17 '清洁运行中'; 18 '换爪位置'; 19 '水平方向钻入位置'; 20 '向上方向钻入位置'; 21 '向下方向钻入位置'; 22 '检查钻头位置'; 23 '请求钻孔'; 24 '请求停止钻孔'; 25 '清洁位置'; 26 '换爪完成'; 27 '水平方向钻入完成'; 28 '向上方向钻入完成'; 29 '向下方向钻入完成'; 30 '检查钻头完成'

text list "DB_PromptStartNotPmt": 1000 '设备不在原点,需要复位!'; 1001 '请摁下自动模式启动按钮！'; 1002 '安全门旁路，注意安全！'; 1003 '安全门电磁线圈锁定失败！'; 1004 '上位机通讯失败！'

text list "DB_PromptBeeper": 2000 '设备紧急停止中,请复位！'; 2001 '设备气压低，请复位！'; 2002 '气源未打开，请摁下复位按钮！'; 2003 '气缸操作条件不满足，请检查！'; 2004 '上位机急停！'; 2005 '打孔超时！'; 2006 '推力缸初始位置不正确！'; 2007 ''; 2008 ''; 2009 '机器人未准备好！'; 2010 '操作盒急停NOK'; 2011 '机器人急停按钮NOK'; 2012 '温控器报警'; 2013 '围栏内侧急停NOK'; 2014 '水泥块击打框架急停NOK'; 2015 ''; 2016 '电源夹具ID号错误，请检查夹具！'; 2017 '低电流工作超时报警！'; 2018 ''; 2019 ''; 2020 ''; 2021 ''; 2022 '光幕被遮，确认安全后复位！'; 2023 '信号夹具ID号错误，请检查夹具！'; 2024 '水平水泥板已打完，请更换水泥板！'; 2025 '垂直向上水泥板已打完，请更换水泥板！'; 2026 '垂直向下水泥板已打完，请更换水泥板！'; 2027 '批头长度错误，请更换！'; 2028 '角度设置超限！'; 2029 '夹具位置已满，无法换型！'; 2030 '钻孔深度超限！'; 2031 '机器人设置速度不能超过100！'; 2032 'Z01.推力气缸工作位置故障!'; 2033 'Z01.推力气缸基本位置故障!'; 2034 'Z02.辅助气缸工作位置故障!'; 2035 'Z02.辅助气缸基本位置故障!'; 2036 'Z03.左防尘盖夹紧缸工作位置故障!'; 2037 'Z03.左防尘盖夹紧缸基本位置故障!'; 2038 'Z04.右防尘盖夹紧缸工作位置故障!'; 2039 'Z04.右防尘盖夹紧缸基本位置故障!'; 2040 'Z05.枪电源工作位置故障!'; 2041 'Z05.枪电源基本位置故障!'; 2042 'Z06.水泥板吹气工作位置故障!'; 2043 'Z06.水泥板吹气基本位置故障!'; 2044 'Z07.快换盘锁紧工作位置故障!'; 2045 'Z07.快换盘锁紧基本位置故障!'; 2046 ''; 2064 ''; 2065 ''; 2066 ''

text list "KuKaRobotStatusPrompt": 0 'A00. ModeOff !'; 1 'A01. OK To Start !'; 2 'A02.Wait User Command = Off!'; 3 'A03.'; 4 'A04. Wait IO.Busy = Off'; 5 'A05. Wait IO.END = ON, Check K3'; 6 'A06. Wait IO.Move = Off, Check K12=?, K23=Move'; 7 'A07. Wait Cmd Ready!'; 8 'A10.'; 9 'A11.'; 10 'A12.'; 11 'A13.'; 12 'A14. Start Change Prog'; 13 'A15. Start Drivers on!'; 14 'A16.Start Ext Start!'; 15 'A17.Start Recovery!'; 16 'A20.Start CmdStart!'; 17 'A21.Wait Done'; 18 'A22.'; 19 'A23.'; 20 'A24.'; 21 'A25.'; 22 'A26.'; 23 'A27.'; 24 'A30.'; 25 'A31'; 26 'A32'; 27 'A33'; 28 'A34'; 29 'A35'; 30 'A36'; 31 'A37.'; 32 'E00. Connnect Err, Pls Reset!'; 33 'E01. Cmd end of time Out !'; 34 'E02. Alarm stop!'; 35 'E03. User Saf!'; 36 'E04. Stop mess!'; 37 'E05.Alarm stop intern!'; 38 'E06.in T1 Mode!'; 39 'E07.in T2 Mode!'; 40 'E10.in AUT Mode!'; 41 'E11.'; 42 'E12.'; 43 'E13.'; 44 'E14.'; 45 'E15'; 46 'E16.'; 47 'E17.'; 48 'E20.'; 49 'E21.'; 50 'E22'; 51 'E23'; 52 'E24'; 53 'E25'; 54 'E26'; 55 'E27'; 56 'E30'; 57 'E31'; 58 'E32'; 59 'E33'; 60 'E34'; 61 'E35'; 62 'E36.'; 63 'E37'

text list "校验": 1 '水平'; 2 '向上'; 3 '向下'

graphic list "语言切换": 0 'Uk'; 1 'China'

screen "01-首页" 1280x1024
   on GenerateScreen: function_bed61462(1)
   on ClearScreen: SetTag("DB_SysMode_TPCurSubPage", 0); SetTag("DB_SysMode_TPCurPageType", 200)
   Button "Button" at 533,426 size 172x123; TextOn '进入'; TextOff '进入'; PictureOn "向右箭头_0"; PictureOff "向右箭头_0"
      on Click: ActivateScreen("200-自动画面", 0)
   TextField "TemplateTextFieldScreenName_0" at 377,594 size 495x31; Text '上海克来机电自动化工程股份有限公司 / 上海克来机电自动化工程有限公司'
   TextField "TemplateTextFieldScreenName_1" at 541,734 size 150x31; Text '2020年10月 / 2013年08月'
   TextField "TemplateTextFieldScreenName_2" at 408,148 size 437x31; Text '杭州博世 / 上海克来机电自动化工程有限公司'
   TextField "TemplateTextFieldScreenName_3" at 406,297 size 437x31; Text '电锤功能测试设备 / 上海克来机电自动化工程有限公司'

screen "09-报警画面" 1280x1024, template "Template"
   Button "按钮_4" at 124,893 size 256x128; TextOn '品种 参数'; TextOff '指示灯测试'
      on Press: function_b14e0dd5("DB_SysMode_TPPB", 0)
      Appearance <- "DB_SysMode_TPPB"
   Button "按钮_6" at 382,893 size 256x128; TextOn '日光灯ON'; TextOff '日光灯'
      on Click: function_c82f6f27("DB_SysMode_TPPB", 4)
      Appearance <- "DB_SysMode_TPPB"
   TextField "文本域_9" at 120,75 size 1040x75; Text '报警信息'
   Button "按钮_1" at 394,252 size 506x171; TextOn '品种 参数'; TextOff '当前报警画面 / 故障复位'
      on Press: ActivateScreen("11-当前报警画面", 0)
   Button "按钮_2" at 394,467 size 506x171; TextOn '品种 参数'; TextOff '历史报警画面 / 故障复位'
      on Press: ActivateScreen("12-历史报警画面", 0)
   Button "按钮_7" at 642,893 size 256x128; TextOn '日光灯ON'; TextOff '蜂鸣器'
      on Click: function_c82f6f27("DB_SysMode_TPPB", 5)
      Appearance <- "DB_SysMode_TPPB"
   Button "按钮_3" at 900,893 size 256x128; TextOn '故障复位 / 日光灯ON'; TextOff '故障复位 / 蜂鸣器'
      on Press: function_b14e0dd5("DB_SysMode_TPPB", 3)
      Appearance <- "DB_SysMode_TPPB"

screen "11-当前报警画面" 1280x1024, template "Template"
   TextField "文本域_11" at 120,75 size 1040x75; Text '当前报警信息 / 报警信息'
   AlarmView "报警视图_1" at 120,149 size 1036x707; ColumnTextDevice 'PLC'; ColumnTextNumber '编号 / No.'; ColumnTextAckGroup 'GR / Acknowledge group'; ColumnTextAlarmState '状态 / Status'; ColumnTextTime '时间 / Time'; ColumnTextDate '日期 / Date'; ColumnTextAlarmText '文本 / Text'
   Button "按钮_5" at 892,868 size 268x141; TextOn '品种 参数'; TextOff '返回 / 故障复位'
      on Press: function_efd93a16()

screen "12-历史报警画面" 1280x1024, template "Template"
   TextField "文本域_12" at 120,75 size 1040x75; Text '历史报警信息 / 报警信息'
   AlarmView "报警视图_1" at 120,149 size 1036x708; ColumnTextDevice 'PLC'; ColumnTextNumber '编号 / No.'; ColumnTextAckGroup 'GR / Acknowledge group'; ColumnTextAlarmState '状态 / Status'; ColumnTextTime '时间 / Time'; ColumnTextDate '日期 / Date'; ColumnTextAlarmText '文本 / Text'
   Button "按钮_5" at 892,869 size 268x141; TextOn '品种 参数'; TextOff '返回 / 故障复位'
      on Press: function_efd93a16()

screen "200-自动画面" 1280x1024, template "Template"
   SymbolicIOField "符号 IO 域_1" at 120,951 size 1040x69; TextOn '1'; TextOff '0'; TextList "操作提示"
      ProcessValue <- "DB_Message_PromptValue"

screen "220-统计信息" 1280x1024, template "Template"
   TextField "文本域_220" at 120,75 size 1040x75; Text '产量统计 / 统计信息'
   SymbolicIOField "符号 IO 域_1" at 120,951 size 1040x69; TextOn '1'; TextOff '0'; TextList "操作提示"
      ProcessValue <- "DB_Message_PromptValue"

screen "240-工位操作" 1280x1024, template "Template"
   TextField "文本域_240" at 120,75 size 1040x75; Text '工位操作 / 校验信息'
   SymbolicIOField "符号 IO 域_1" at 120,951 size 1040x69; TextOn '1'; TextOff '0'; TextList "操作提示"
      ProcessValue <- "DB_Message_PromptValue"
   Button "按钮_21" at 232,269 size 272x192; TextOff '单工位自动'
      on Press: ActivateScreen("241-单工位自动", 0)
   Button "按钮_1" at 508,269 size 272x192; TextOff '单工位回原点'
      on Press: ActivateScreen("242-单工位回原点", 0)
   Button "按钮_2" at 782,269 size 272x192; TextOff '...'
   Button "按钮_3" at 232,467 size 272x192; TextOff '...'
   Button "按钮_4" at 508,467 size 272x192; TextOff '...'
   Button "按钮_5" at 782,467 size 272x192; TextOff '...'
   Button "按钮_6" at 232,661 size 272x192; TextOff '...'
   Button "按钮_7" at 508,661 size 272x192; TextOff '...'
   Button "按钮_8" at 782,661 size 272x192; TextOff '...'

screen "241-单工位自动" 1280x1024, template "Template"
   TextField "文本域_200" at 120,75 size 1040x75; Text '单工位自动 / 自动操作'
   SymbolicIOField "符号 IO 域_1" at 120,951 size 1040x69; TextOn '1'; TextOff '0'; TextList "操作提示"
      ProcessValue <- "DB_Message_PromptValue"
   Button "按钮_21" at 154,157 size 260x147; TextOff '01.托盘上料 启动 ******* 基本位Z1'
   Button "按钮_1" at 154,317 size 260x147; TextOff 'xxxx启动 ******* 基本位Z1'
   Button "按钮_2" at 154,476 size 260x147; TextOff 'xxxx启动 ******* 基本位Z1'
   Button "按钮_3" at 154,635 size 260x147; TextOff 'xxxx启动 ******* 基本位Z1'
   Button "按钮_4" at 154,791 size 260x147; TextOff 'xxxx启动 ******* 基本位Z1'
   Button "按钮_5" at 486,157 size 266x147; TextOff 'xxxx启动 ******* 基本位Z1'
   Button "按钮_6" at 486,316 size 266x147; TextOff 'xxxx启动 ******* 基本位Z1'
   Button "按钮_7" at 486,476 size 266x147; TextOff 'xxxx启动 ******* 基本位Z1'
   Button "按钮_8" at 486,635 size 262x147; TextOff 'xxxx启动 ******* 基本位Z1'
   Button "按钮_9" at 820,157 size 262x147; TextOff 'xxxx启动 ******* 基本位Z1'
   Button "按钮_10" at 820,476 size 262x147; TextOff 'xxxx启动 ******* 基本位Z1'
   Button "按钮_11" at 820,635 size 262x147; TextOff 'xxxx启动 ******* 基本位Z1'
   Button "按钮_12" at 820,315 size 262x147; TextOff 'xxxx启动 ******* 基本位Z1'
   Button "按钮_13" at 1022,841 size 128x96; TextOn '品种 参数'; TextOff '返回 / 故障复位'
      on Press: function_efd93a16()

screen "242-单工位回原点" 1280x1024, template "Template"
   TextField "文本域_241" at 120,75 size 1040x75; Text '单工位回原点 / 校验信息'
   SymbolicIOField "符号 IO 域_1" at 120,949 size 1040x69; TextOn '1'; TextOff '0'; TextList "操作提示"
      ProcessValue <- "DB_Message_PromptValue"
   Button "按钮_6" at 244,403 size 310x183; TextOff 'xxx工位回原点 ******* 基本位Z1'
   Button "按钮_7" at 244,621 size 310x181; TextOff 'xxx工位回原点 ******* 基本位Z1'
   Button "按钮_9" at 666,188 size 308x181; TextOff 'xxx工位回原点 ******* 基本位Z1'
   Button "按钮_12" at 666,403 size 308x181; TextOff 'xxx工位回原点 ******* 基本位Z1'
   Button "按钮_13" at 1022,841 size 128x96; TextOn '品种 参数'; TextOff '返回 / 故障复位'
      on Press: function_efd93a16()

screen "201-特殊模式" 1280x1024, template "Template"
   TextField "文本域_140" at 120,75 size 1040x75; Text '特殊模式选择 / 伺服点动'
   SymbolicIOField "符号 IO 域_1" at 120,951 size 1040x69; TextOn '1'; TextOff '0'; TextList "操作提示"
      ProcessValue <- "DB_Message_PromptValue"
   Button "按钮_9" at 914,891 size 244x123; TextOff '返 回'
      on Press: function_efd93a16()
   Button "按钮_21" at 232,269 size 272x192; TextOff '单步调试'
      on Press: function_c82f6f27("DB_SysMode_TPPB", 2)
      Appearance <- "DB_SysMode_TPPB"
   Button "按钮_1" at 508,269 size 272x192; TextOff '...'
   Button "按钮_2" at 782,269 size 272x192; TextOff '...'
   Button "按钮_3" at 232,467 size 272x192; TextOff '...'
   Button "按钮_4" at 508,467 size 272x192; TextOff '...'
   Button "按钮_5" at 782,467 size 272x192; TextOff '...'
   Button "按钮_6" at 232,661 size 272x192; TextOff '...'
   Button "按钮_7" at 508,661 size 272x192; TextOff '...'
   Button "按钮_8" at 782,661 size 272x192; TextOff '临时屏蔽设定'
      on Press: ActivateScreen("209-临时屏蔽", 0)
      Appearance <- "DB_SysMode_DisableOption"

screen "209-临时屏蔽" 1280x1024, template "Template"
   TextField "文本域_140" at 120,75 size 1040x75; Text '临时屏蔽选项 / 伺服点动'
   SymbolicIOField "符号 IO 域_1" at 118,949 size 1040x69; TextOn '1'; TextOff '0'; TextList "操作提示"
      ProcessValue <- "DB_Message_PromptValue"
   Button "按钮_9" at 914,891 size 244x123; TextOff '返 回'
      on Press: function_efd93a16()
   Button "按钮_21" at 132,179 size 252x139; TextOff 'xx相机屏蔽'
      on Press: function_c82f6f27("DB_SysMode_DisableOption", 8)
      Appearance <- "DB_SysMode_DisableOption"
   Button "按钮_1" at 388,179 size 252x139; TextOff '屏蔽项-2'
      on Press: function_c82f6f27("DB_SysMode_DisableOption", 9)
      Appearance <- "DB_SysMode_DisableOption"
   Button "按钮_2" at 644,179 size 252x139; TextOff '...'
      on Press: function_c82f6f27("DB_SysMode_DisableOption", 10)
      Appearance <- "DB_SysMode_DisableOption"
   Button "按钮_3" at 132,329 size 252x139; TextOff '...'
      on Press: function_c82f6f27("DB_SysMode_DisableOption", 12)
      Appearance <- "DB_SysMode_DisableOption"
   Button "按钮_4" at 388,329 size 252x139; TextOff '...'
      on Press: function_c82f6f27("DB_SysMode_DisableOption", 13)
      Appearance <- "DB_SysMode_DisableOption"
   Button "按钮_5" at 644,329 size 252x139; TextOff '...'
      on Press: function_c82f6f27("DB_SysMode_DisableOption", 14)
      Appearance <- "DB_SysMode_DisableOption"
   Button "按钮_6" at 132,483 size 252x139; TextOff '...'
      on Press: function_c82f6f27("DB_SysMode_DisableOption", 0)
      Appearance <- "DB_SysMode_DisableOption"
   Button "按钮_7" at 388,483 size 252x139; TextOff '...'
      on Press: function_c82f6f27("DB_SysMode_DisableOption", 1)
      Appearance <- "DB_SysMode_DisableOption"
   Button "按钮_8" at 644,483 size 252x139; TextOff '...'
      on Press: function_c82f6f27("DB_SysMode_DisableOption", 2)
      Appearance <- "DB_SysMode_DisableOption"
   Button "按钮_10" at 900,179 size 252x139; TextOff '...'
      on Press: function_c82f6f27("DB_SysMode_DisableOption", 11)
      Appearance <- "DB_SysMode_DisableOption"
   Button "按钮_11" at 900,329 size 252x139; TextOff '...'
      on Press: function_c82f6f27("DB_SysMode_DisableOption", 15)
      Appearance <- "DB_SysMode_DisableOption"
   Button "按钮_12" at 900,483 size 252x139; TextOff '...'
      on Press: function_c82f6f27("DB_SysMode_DisableOption", 3)
      Appearance <- "DB_SysMode_DisableOption"
   Button "按钮_13" at 132,636 size 252x139; TextOff '...'
      on Press: function_c82f6f27("DB_SysMode_DisableOption", 4)
      Appearance <- "DB_SysMode_DisableOption"
   Button "按钮_14" at 388,636 size 252x139; TextOff '...'
      on Press: function_c82f6f27("DB_SysMode_DisableOption", 5)
      Appearance <- "DB_SysMode_DisableOption"
   Button "按钮_15" at 644,636 size 252x139; TextOff '...'
      on Press: function_c82f6f27("DB_SysMode_DisableOption", 6)
      Appearance <- "DB_SysMode_DisableOption"
   Button "按钮_16" at 900,636 size 252x139; TextOff '...'
      on Press: function_c82f6f27("DB_SysMode_DisableOption", 7)
      Appearance <- "DB_SysMode_DisableOption"

screen "260- IO_Check主页面" 1280x1024, template "Template"
   TextField "文本域_260" at 120,75 size 1040x75; Text 'IO状态查看'
   SymbolicIOField "符号 IO 域_1" at 123,951 size 1040x64; TextOn '1'; TextOff '0'; TextList "操作提示"
      ProcessValue <- "DB_Message_PromptValue"
   Button "按钮_21" at 232,269 size 272x192; TextOff '常规IO I0.0-I9.7 Q0.0-Q5.7'
      on Release: ActivateScreen("261_IOCheck_Input", 0)
      on Press: SetTag("DB_IOCheck____InputMinByteNo", 0); SetTag("DB_IOCheck____InputMaxByteNo", 9); SetTag("DB_IOCheck____OutputMinByteNo", 0); SetTag("DB_IOCheck____OutputMaxByteNo", 5)
   Button "按钮_2" at 507,269 size 272x192; TextOff '阀岛IO I20.0-I31.7 Q20.0-Q29.7'
      on Release: ActivateScreen("261_IOCheck_Input", 0)
      on Press: SetTag("DB_IOCheck____InputMinByteNo", 20); SetTag("DB_IOCheck____InputMaxByteNo", 31); SetTag("DB_IOCheck____OutputMinByteNo", 20); SetTag("DB_IOCheck____OutputMaxByteNo", 29)
   Button "按钮_3" at 782,269 size 272x192; TextOff '阀岛IO I36.0-I43.7 Q30.0-Q38.7'
      on Release: ActivateScreen("261_IOCheck_Input", 0)
      on Press: SetTag("DB_IOCheck____InputMinByteNo", 36); SetTag("DB_IOCheck____InputMaxByteNo", 43); SetTag("DB_IOCheck____OutputMinByteNo", 30); SetTag("DB_IOCheck____OutputMaxByteNo", 38)
   Button "按钮_5" at 232,465 size 272x192; TextOff '...'
      on Release: ActivateScreen("261_IOCheck_Input", 0)
      on Press: SetTag("DB_IOCheck____InputMinByteNo", 20); SetTag("DB_IOCheck____InputMaxByteNo", 35); SetTag("DB_IOCheck____OutputMinByteNo", 20); SetTag("DB_IOCheck____OutputMaxByteNo", 30)
   Button "按钮_6" at 507,465 size 272x192; TextOff '...'
      on Release: ActivateScreen("261_IOCheck_Input", 0)
      on Press: SetTag("DB_IOCheck____InputMinByteNo", 20); SetTag("DB_IOCheck____InputMaxByteNo", 35); SetTag("DB_IOCheck____OutputMinByteNo", 20); SetTag("DB_IOCheck____OutputMaxByteNo", 30)
   Button "按钮_7" at 782,465 size 272x192; TextOff '...'
      on Release: ActivateScreen("261_IOCheck_Input", 0)
      on Press: SetTag("DB_IOCheck____InputMinByteNo", 20); SetTag("DB_IOCheck____InputMaxByteNo", 35); SetTag("DB_IOCheck____OutputMinByteNo", 20); SetTag("DB_IOCheck____OutputMaxByteNo", 30)
   Button "按钮_8" at 232,661 size 272x192; TextOff '...'
      on Release: ActivateScreen("261_IOCheck_Input", 0)
      on Press: SetTag("DB_IOCheck____InputMinByteNo", 20); SetTag("DB_IOCheck____InputMaxByteNo", 35); SetTag("DB_IOCheck____OutputMinByteNo", 20); SetTag("DB_IOCheck____OutputMaxByteNo", 30)
   Button "按钮_9" at 507,661 size 272x192; TextOff '...'
      on Release: ActivateScreen("261_IOCheck_Input", 0)
      on Press: SetTag("DB_IOCheck____InputMinByteNo", 20); SetTag("DB_IOCheck____InputMaxByteNo", 35); SetTag("DB_IOCheck____OutputMinByteNo", 20); SetTag("DB_IOCheck____OutputMaxByteNo", 30)
   Button "按钮_10" at 782,661 size 272x192; TextOff '...'
      on Release: ActivateScreen("261_IOCheck_Input", 0)
      on Press: SetTag("DB_IOCheck____InputMinByteNo", 20); SetTag("DB_IOCheck____InputMaxByteNo", 35); SetTag("DB_IOCheck____OutputMinByteNo", 20); SetTag("DB_IOCheck____OutputMaxByteNo", 30)

screen "261_IOCheck_Input" 1280x1024, template "Template"
   SymbolicIOField "符号 IO 域_1" at 125,160 size 203x77; TextOn '1'; TextOff '0'; TextList "Input_地址"
      ProcessValue <- "[0]"
      Appearance <- "IO_Input_SignalStatus"
   SymbolicIOField "符号 IO 域_2" at 333,160 size 819x77; TextOn '1'; TextOff '0'; TextList "Input_注释"
      ProcessValue <- "[0]"
   SymbolicIOField "符号 IO 域_31" at 125,243 size 203x77; TextOn '1'; TextOff '0'; TextList "Input_地址"
      ProcessValue <- "[1]"
      Appearance <- "IO_Input_SignalStatus"
   SymbolicIOField "符号 IO 域_32" at 333,243 size 819x77; TextOn '1'; TextOff '0'; TextList "Input_注释"
      ProcessValue <- "[1]"
   SymbolicIOField "符号 IO 域_33" at 125,322 size 203x75; TextOn '1'; TextOff '0'; TextList "Input_地址"
      ProcessValue <- "[2]"
      Appearance <- "IO_Input_SignalStatus"
   SymbolicIOField "符号 IO 域_34" at 333,322 size 819x75; TextOn '1'; TextOff '0'; TextList "Input_注释"
      ProcessValue <- "[2]"
   SymbolicIOField "符号 IO 域_35" at 125,405 size 203x75; TextOn '1'; TextOff '0'; TextList "Input_地址"
      ProcessValue <- "[3]"
      Appearance <- "IO_Input_SignalStatus"
   SymbolicIOField "符号 IO 域_36" at 333,403 size 819x77; TextOn '1'; TextOff '0'; TextList "Input_注释"
      ProcessValue <- "[3]"
   SymbolicIOField "符号 IO 域_37" at 125,495 size 203x81; TextOn '1'; TextOff '0'; TextList "Input_地址"
      ProcessValue <- "[4]"
      Appearance <- "IO_Input_SignalStatus"
   SymbolicIOField "符号 IO 域_38" at 333,495 size 819x81; TextOn '1'; TextOff '0'; TextList "Input_注释"
      ProcessValue <- "[4]"
   SymbolicIOField "符号 IO 域_39" at 125,578 size 203x79; TextOn '1'; TextOff '0'; TextList "Input_地址"
      ProcessValue <- "[5]"
      Appearance <- "IO_Input_SignalStatus"
   SymbolicIOField "符号 IO 域_40" at 333,578 size 819x79; TextOn '1'; TextOff '0'; TextList "Input_注释"
      ProcessValue <- "[5]"
   SymbolicIOField "符号 IO 域_41" at 125,661 size 203x75; TextOn '1'; TextOff '0'; TextList "Input_地址"
      ProcessValue <- "[6]"
      Appearance <- "IO_Input_SignalStatus"
   SymbolicIOField "符号 IO 域_42" at 333,661 size 819x75; TextOn '1'; TextOff '0'; TextList "Input_注释"
      ProcessValue <- "[6]"
   SymbolicIOField "符号 IO 域_43" at 125,745 size 203x77; TextOn '1'; TextOff '0'; TextList "Input_地址"
      ProcessValue <- "[7]"
      Appearance <- "IO_Input_SignalStatus"
   SymbolicIOField "符号 IO 域_44" at 333,745 size 819x77; TextOn '1'; TextOff '0'; TextList "Input_注释"
      ProcessValue <- "[7]"
   TextField "文本域_261" at 384,75 size 552x85; Text 'InPut状态'
   Button "按钮_4" at 125,881 size 208x130; TextOff '<<'
      on Press: function_b9b71300("DB_IOCheck____In_ByteNo", 1)
      Appearance <- "DB_IOCheck____TP_Status"
      ObjectEnable <- "DB_IOCheck____TP_Status"
   Button "按钮_5" at 693,881 size 211x130; TextOff '>>'
      on Press: function_dd21b452("DB_IOCheck____In_ByteNo", 1)
      Appearance <- "DB_IOCheck____TP_Status"
      ObjectEnable <- "DB_IOCheck____TP_Status"
   Button "按钮_6" at 381,881 size 264x130; TextOff '->OutPut'
      on Release: ActivateScreen("262_IOCheck_Output", 0)
   Button "按钮_7" at 936,881 size 216x130; TextOff '返回'
      on Click: ActivateScreen("260- IO_Check主页面", 0)

screen "262_IOCheck_Output" 1280x1024, template "Template"
   SymbolicIOField "符号 IO 域_1" at 125,160 size 203x79; TextOn '1'; TextOff '0'; TextList "OutPut_地址"
      ProcessValue <- "[0]"
      Appearance <- "IO_OutPut_SignalStatus"
   SymbolicIOField "符号 IO 域_2" at 337,161 size 819x79; TextOn '1'; TextOff '0'; TextList "OutPut_注释"
      ProcessValue <- "[0]"
   SymbolicIOField "符号 IO 域_31" at 125,243 size 203x77; TextOn '1'; TextOff '0'; TextList "OutPut_地址"
      ProcessValue <- "[1]"
      Appearance <- "IO_OutPut_SignalStatus"
   SymbolicIOField "符号 IO 域_32" at 337,244 size 819x77; TextOn '1'; TextOff '0'; TextList "OutPut_注释"
      ProcessValue <- "[1]"
   SymbolicIOField "符号 IO 域_33" at 125,324 size 203x75; TextOn '1'; TextOff '0'; TextList "OutPut_地址"
      ProcessValue <- "[2]"
      Appearance <- "IO_OutPut_SignalStatus"
   SymbolicIOField "符号 IO 域_34" at 337,325 size 819x75; TextOn '1'; TextOff '0'; TextList "OutPut_注释"
      ProcessValue <- "[2]"
   SymbolicIOField "符号 IO 域_35" at 125,403 size 203x77; TextOn '1'; TextOff '0'; TextList "OutPut_地址"
      ProcessValue <- "[3]"
      Appearance <- "IO_OutPut_SignalStatus"
   SymbolicIOField "符号 IO 域_36" at 337,404 size 819x77; TextOn '1'; TextOff '0'; TextList "OutPut_注释"
      ProcessValue <- "[3]"
   SymbolicIOField "符号 IO 域_37" at 125,497 size 203x77; TextOn '1'; TextOff '0'; TextList "OutPut_地址"
      ProcessValue <- "[4]"
      Appearance <- "IO_OutPut_SignalStatus"
   SymbolicIOField "符号 IO 域_38" at 333,660 size 819x77; TextOn '1'; TextOff '0'; TextList "OutPut_注释"
      ProcessValue <- "[6]"
   SymbolicIOField "符号 IO 域_39" at 125,578 size 203x79; TextOn '1'; TextOff '0'; TextList "OutPut_地址"
      ProcessValue <- "[5]"
      Appearance <- "IO_OutPut_SignalStatus"
   SymbolicIOField "符号 IO 域_40" at 333,497 size 819x79; TextOn '1'; TextOff '0'; TextList "OutPut_注释"
      ProcessValue <- "[4]"
   SymbolicIOField "符号 IO 域_41" at 125,659 size 203x79; TextOn '1'; TextOff '0'; TextList "OutPut_地址"
      ProcessValue <- "[6]"
      Appearance <- "IO_OutPut_SignalStatus"
   SymbolicIOField "符号 IO 域_42" at 333,577 size 819x79; TextOn '1'; TextOff '0'; TextList "OutPut_注释"
      ProcessValue <- "[5]"
   SymbolicIOField "符号 IO 域_43" at 125,742 size 203x77; TextOn '1'; TextOff '0'; TextList "OutPut_地址"
      ProcessValue <- "[7]"
      Appearance <- "IO_OutPut_SignalStatus"
   SymbolicIOField "符号 IO 域_44" at 333,741 size 819x77; TextOn '1'; TextOff '0'; TextList "OutPut_注释"
      ProcessValue <- "[7]"
   TextField "OutPut" at 384,75 size 552x85; Text 'OutPut状态'
   Button "按钮_4" at 125,881 size 208x128; TextOff '<<'
      on Press: function_b9b71300("DB_IOCheck____Out_ByteNo", 1)
      Appearance <- "DB_IOCheck____TP_Status"
      ObjectEnable <- "DB_IOCheck____TP_Status"
   Button "按钮_5" at 693,881 size 211x128; TextOff '>>'
      on Press: function_dd21b452("DB_IOCheck____Out_ByteNo", 1)
      Appearance <- "DB_IOCheck____TP_Status"
      ObjectEnable <- "DB_IOCheck____TP_Status"
   Button "按钮_6" at 381,881 size 264x128; TextOff 'InPut<-'
      on Release: ActivateScreen("261_IOCheck_Input", 0)
   Button "按钮_7" at 936,881 size 216x128; TextOff '返回'
      on Click: ActivateScreen("260- IO_Check主页面", 0)

screen "380-主画面" 1280x1024, template "Template"
   TextField "仪器程序号" at 120,75 size 1040x75; Text '系统设定选择 / 仪器程序号'
   IOField "IO 域_28" at 380,883 size 108x128; FormatPattern 99
      ProcessValue <- "DB_Parameter_CurProgNoE"
   TextField "文本域_2" at 120,892 size 112x115; Text '型号 选择：'
   IOField "IO 域_2" at 496,883 size 308x128; FormatPattern ?????????????
      ProcessValue <- "DB_Parameter_TypeParaE_TypeName"
   Button "按钮_4" at 232,883 size 140x132; TextOff '<<'
      on Press: function_b9b71300("DB_Parameter_CurProgNoE", 1)
      ObjectEnable <- "DB_Parameter_CurProgNoE"
   Button "按钮_5" at 812,883 size 140x132; TextOff '>>'
      on Press: function_dd21b452("DB_Parameter_CurProgNoE", 1)
      ObjectEnable <- "DB_Parameter_CurProgNoE"
   Button "按钮_3" at 965,883 size 188x132; TextOff '保 存'
      on Press: function_b14e0dd5("DB_Parameter_TP_Cmd", 8)
      Appearance <- "DB_Parameter_TP_Status"
   Button "按钮_21" at 232,224 size 272x192; TextOff '01.X轴伺服 参数'
      on Press: ActivateScreen("301-时间设置", 0)
   Button "按钮_1" at 508,224 size 272x192; TextOff '...'
      on Press: ActivateScreen("301-时间设置", 0)
   Button "按钮_2" at 782,224 size 272x192; TextOff '...'
      on Press: ActivateScreen("301-时间设置", 0)
   Button "按钮_6" at 232,420 size 272x192; TextOff '...'
      on Press: ActivateScreen("301-时间设置", 0)
   Button "按钮_7" at 508,420 size 272x192; TextOff '...'
      on Press: ActivateScreen("301-时间设置", 0)
   Button "按钮_8" at 782,420 size 272x192; TextOff '...'
      on Press: ActivateScreen("301-时间设置", 0)
   Button "按钮_9" at 232,617 size 272x192; TextOff '...'
      on Press: ActivateScreen("301-时间设置", 0)
   Button "按钮_10" at 508,617 size 272x192; TextOff '用户权限 管理'
      on Press: ActivateScreen("388-用户管理", 0)
   Button "按钮_11" at 782,617 size 272x192; TextOff '时间设置'
      on Press: ActivateScreen("389-时间设置", 0)

screen "381-设定1" 1280x1024, template "Template"
   TextField "文本域_601" at 120,75 size 1040x75; Text '系统参数 / 仪器程序号'
   Button "按钮_3" at 906,891 size 244x123; TextOff '返 回'
      on Press: ActivateScreen("360-xxx", 0)
   TextField "文本域_113" at 130,157 size 218x75; Text '当前时间: / 仪器程序号'
   TextField "文本域_114" at 130,237 size 218x75; Text '设定时间: / 仪器程序号'
   Button "按钮_8" at 656,891 size 244x123; TextOff '保 存'
      on Press: function_b14e0dd5("DB_Parameter_TP_Cmd", 8)
      Appearance <- "DB_Parameter_TP_Status"
   DateTimeField "日期/时间域_1" at 352,237 size 295x31
      ProcessValue <- "DB_SysMode_Sys_Time_SetPLCTimeTP"
   DateTimeField "日期/时间域_2" at 352,155 size 295x31
      ProcessValue <- "DB_SysMode_Sys_Time_CurPLCTime"

screen "389-时间设置" 1280x1024, template "Template"
   TextField "文本域_602" at 120,75 size 1040x75; Text '时间设置 / 仪器程序号'
   TextField "文本域_113" at 130,157 size 218x75; Text '当前时间: / 仪器程序号'
   TextField "文本域_114" at 130,237 size 218x75; Text '设定时间: / 仪器程序号'
   Button "按钮_3" at 908,887 size 244x123; TextOff '返 回'
      on Press: ActivateScreen("360-xxx", 0)
   DateTimeField "日期/时间域_1" at 352,237 size 295x31
      ProcessValue <- "DB_SysMode_Sys_Time_SetPLCTimeTP"
   DateTimeField "日期/时间域_2" at 352,155 size 295x31
      ProcessValue <- "DB_SysMode_Sys_Time_CurPLCTime"

screen "388-用户管理" 1280x1024, template "Template"
   UserView "UserView" at 124,160 size 1028x693
   TextField "文本域_5" at 120,73 size 1040x77; Text '用户管理'
   Button "按钮_3" at 908,887 size 244x123; TextOff '返 回'
      on Press: ActivateScreen("360-xxx", 0)

screen "300-主页面" 1280x1024, template "Template"
   TextField "仪器程序号" at 120,75 size 1040x75; Text '系统参数 / 仪器程序号'
   IOField "IO 域_28" at 380,883 size 108x128; FormatPattern 99
      ProcessValue <- "DB_Parameter_CurProgNoE"
   TextField "文本域_2" at 120,892 size 112x115; Text '型号 选择：'
   IOField "IO 域_2" at 496,883 size 308x128; FormatPattern ?????????????
      ProcessValue <- "DB_Parameter_TypeParaE_TypeName"
   Button "按钮_4" at 232,883 size 140x132; TextOff '<<'
      on Press: function_b9b71300("DB_Parameter_CurProgNoE", 1)
      ObjectEnable <- "DB_Parameter_CurProgNoE"
   Button "按钮_5" at 812,883 size 140x132; TextOff '>>'
      on Press: function_dd21b452("DB_Parameter_CurProgNoE", 1)
      ObjectEnable <- "DB_Parameter_CurProgNoE"
   Button "按钮_3" at 952,883 size 201x130; TextOff '保 存'
      on Press: function_b14e0dd5("DB_Parameter_TP_Cmd", 8)
      Appearance <- "DB_Parameter_TP_Status"

screen "301-时间设置" 1280x1024, template "Template"
   TextField "左侧平移伺服参数" at 120,75 size 1040x75; Text '时间设置 / 仪器程序号'
   IOField "IO 域_28" at 380,883 size 108x128; FormatPattern 99
      ProcessValue <- "DB_Parameter_CurProgNoE"
   TextField "文本域_2" at 120,892 size 112x115; Text '型号 选择：'
   IOField "IO 域_2" at 496,883 size 308x128; FormatPattern ?????????????
      ProcessValue <- "DB_Parameter_TypeParaE_TypeName"
   Button "按钮_4" at 232,883 size 140x132; TextOff '<<'
      on Press: function_b9b71300("DB_Parameter_CurProgNoE", 1)
      ObjectEnable <- "DB_Parameter_CurProgNoE"
   Button "按钮_5" at 812,883 size 140x132; TextOff '>>'
      on Press: function_dd21b452("DB_Parameter_CurProgNoE", 1)
      ObjectEnable <- "DB_Parameter_CurProgNoE"
   IOField "I/O 域_1" at 224,170 size 96x40; FormatPattern 99999
      ProcessValue <- "DB_Component_Aux_SysTimeSet_YEAR"
   TextField "文本域" at 175,175 size 57x29; Text '年'
   IOField "I/O 域_2" at 224,219 size 96x40; FormatPattern 999
      ProcessValue <- "DB_Component_Aux_SysTimeSet_MONTH"
   TextField "文本域_3" at 174,224 size 57x29; Text '月'

screen "320-xxx" 1280x1024, template "Template"
   TextField "文本域_320" at 120,75 size 1040x75; Text '夹具编码 / 仪器程序号'
   IOField "IO 域_28" at 380,883 size 108x128; FormatPattern 99
      ProcessValue <- "DB_Parameter_CurProgNoE"
   TextField "文本域_2" at 120,892 size 112x115; Text '型号 选择：'
   IOField "IO 域_2" at 496,883 size 308x128; FormatPattern ?????????????
      ProcessValue <- "DB_Parameter_TypeParaE_TypeName"
   Button "按钮_4" at 232,883 size 140x132; TextOff '<<'
      on Press: function_b9b71300("DB_Parameter_CurProgNoE", 1)
      ObjectEnable <- "DB_Parameter_CurProgNoE"
   Button "按钮_5" at 812,883 size 140x132; TextOff '>>'
      on Press: function_dd21b452("DB_Parameter_CurProgNoE", 1)
      ObjectEnable <- "DB_Parameter_CurProgNoE"

screen "340-xxx" 1280x1024, template "Template"
   TextField "文本域_340" at 120,75 size 1040x75; Text '仪器程序号'
   IOField "IO 域_28" at 380,883 size 108x128; FormatPattern 99
      ProcessValue <- "DB_Parameter_CurProgNoE"
   TextField "文本域_2" at 120,892 size 112x115; Text '型号 选择：'
   IOField "IO 域_2" at 496,883 size 308x128; FormatPattern ?????????????
      ProcessValue <- "DB_Parameter_TypeParaE_TypeName"
   Button "按钮_4" at 232,883 size 140x132; TextOff '<<'
      on Press: function_b9b71300("DB_Parameter_CurProgNoE", 1)
      ObjectEnable <- "DB_Parameter_CurProgNoE"
   Button "按钮_5" at 812,883 size 140x132; TextOff '>>'
      on Press: function_dd21b452("DB_Parameter_CurProgNoE", 1)
      ObjectEnable <- "DB_Parameter_CurProgNoE"
   TextField "文本域_3" at 132,173 size 112x23; Text '01.xxxxxx:'

screen "360-xxx" 1280x1024, template "Template"
   TextField "文本域_360" at 120,75 size 1040x75; Text '系统参数设定 / 系统参数设定...'
   IOField "IO 域_28" at 380,883 size 108x128; FormatPattern 99
      ProcessValue <- "DB_Parameter_CurProgNoE"
   TextField "文本域_2" at 120,892 size 112x115; Text '型号 选择：'
   IOField "IO 域_2" at 496,883 size 308x128; FormatPattern ?????????????
      ProcessValue <- "DB_Parameter_TypeParaE_TypeName"
   Button "按钮_4" at 232,883 size 140x132; TextOff '<<'
      on Press: function_b9b71300("DB_Parameter_CurProgNoE", 1)
      ObjectEnable <- "DB_Parameter_CurProgNoE"
   Button "按钮_5" at 812,883 size 140x132; TextOff '>>'
      on Press: function_dd21b452("DB_Parameter_CurProgNoE", 1)
      ObjectEnable <- "DB_Parameter_CurProgNoE"
   Button "按钮_2" at 416,277 size 472x183; TextOff '系统参数设定'
      on Press: ActivateScreen("381-设定1", 0)

screen "120-主页面****************" 1280x1024, template "Template"
   TextField "文本域_120" at 120,75 size 1040x75; Text '自动操作'
   SymbolicIOField "符号 IO 域_1" at 120,951 size 1040x69; TextOn '1'; TextOff '0'; TextList "操作提示"
      ProcessValue <- "DB_Message_PromptValue"
   Button "按钮_21" at 232,269 size 272x192; TextOff '...'
   Button "按钮_1" at 508,269 size 272x192; TextOff '...'
   Button "按钮_2" at 782,269 size 272x192; TextOff '...'
   Button "按钮_3" at 232,467 size 272x192; TextOff '...'
   Button "按钮_4" at 508,467 size 272x192; TextOff '...'
   Button "按钮_5" at 782,467 size 272x192; TextOff '...'
   Button "按钮_6" at 232,661 size 272x192; TextOff '...'
   Button "按钮_7" at 508,661 size 272x192; TextOff '...'
   Button "按钮_8" at 782,661 size 272x192; TextOff '...'

screen "140-主页面****************" 1280x1024, template "Template"
   TextField "文本域_140" at 120,75 size 1040x75; Text '测试页面 / 伺服点动'
   SymbolicIOField "符号 IO 域_1" at 120,951 size 1040x69; TextOn '1'; TextOff '0'; TextList "操作提示"
      ProcessValue <- "DB_Message_PromptValue"
   Button "按钮_21" at 232,269 size 272x192; TextOff '...'
   Button "按钮_1" at 508,269 size 272x192; TextOff '...'
   Button "按钮_2" at 782,269 size 272x192; TextOff '...'
   Button "按钮_3" at 232,467 size 272x192; TextOff '...'
   Button "按钮_4" at 508,467 size 272x192; TextOff '...'
   Button "按钮_5" at 782,467 size 272x192; TextOff '...'
   Button "按钮_6" at 232,661 size 272x192; TextOff '...'
   Button "按钮_7" at 508,661 size 272x192; TextOff '...'
   Button "按钮_8" at 782,661 size 272x192; TextOff '...'

screen "160-主页面" 1280x1024, template "Template"
   TextField "文本域_140" at 120,75 size 1040x75; Text 'Laser Mark / 伺服点动'
   SymbolicIOField "符号 IO 域_1" at 118,949 size 1040x69; TextOn '1'; TextOff '0'; TextList "操作提示"
      ProcessValue <- "DB_Message_PromptValue"
   Button "按钮_1" at 508,269 size 272x192; TextOff '...'
   Button "按钮_2" at 782,269 size 272x192; TextOff '...'
   Button "按钮_3" at 232,467 size 272x192; TextOff '...'
   Button "按钮_4" at 508,467 size 272x192; TextOff '...'
   Button "按钮_5" at 782,467 size 272x192; TextOff '...'
   Button "按钮_6" at 232,661 size 272x192; TextOff '...'
   Button "按钮_7" at 508,661 size 272x192; TextOff '...'
   Button "按钮_8" at 782,661 size 272x192; TextOff '...'

screen "190-气缸控制" 1280x1024
   Button "模板_按钮_23" at 1160,0 size 120x192; TextOn '运行 设置'; TextOff '上 页'
      on Press: function_dbe01993("DB_SysMode_Cylinder_Index", 1, "DB_SysMode_Cylinder_Index", -5)
   Button "模板_按钮_24" at 1160,621 size 120x192; TextOn '运行 设置'; TextOff '下 页'
      on Press: function_dbe01993("DB_SysMode_Cylinder_Index", 1, "DB_SysMode_Cylinder_Index", 5)
   Button "模板_按钮_25" at 1160,211 size 120x192; TextOn '运行 设置'; TextOff '+1'; PictureOff "向上箭头"
      on Press: function_dbe01993("DB_SysMode_Cylinder_Index", 1, "DB_SysMode_Cylinder_Index", -1)
   Button "模板_按钮_26" at 1160,416 size 120x192; TextOn '运行 设置'; TextOff '+1'; PictureOff "向下箭头"
      on Press: function_dbe01993("DB_SysMode_Cylinder_Index", 1, "DB_SysMode_Cylinder_Index", 1)
   Button "模板_按钮_33" at 1160,827 size 120x192; TextOn '运行 设置'; TextOff '返回 自动 监视'
      on Click: function_efd93a16()
   SymbolicIOField "符号 IO 域_1" at 0,950 size 1158x69; TextOn '1'; TextOff '0'; TextList "操作提示"
      ProcessValue <- "DB_Message_PromptValue"
   Group "Group" at 12,19 size 1138x921
   Button "按钮_14" at 720,205 size 200x163; TextOff '工作位'
      on Press: function_b14e0dd5("Z02_CmdW", 0)
      Appearance <- "Z02_Status"
   Button "按钮_20" at 12,205 size 468x163; TextOff '******* 基本位Z1'; TextList "Cylinder_Name"
      on Press: function_b14e0dd5("Z02_CmdW", 1)
      Appearance <- "Z02_Status"
      ProcessValue <- "手动控制\CylinderIndex2"
   SymbolicIOField "符号 IO 域_6" at 546,285 size 164x83; TextOn '1'; TextOff '0'; TextList "Cylinder_QRet"
      ProcessValue <- "手动控制\CylinderIndex2"
      Appearance <- "Z02_Status"
   SymbolicIOField "符号 IO 域_7" at 986,285 size 164x83; TextOn '1'; TextOff '0'; TextList "Cylinder_QExt"
      ProcessValue <- "手动控制\CylinderIndex2"
      Appearance <- "Z02_Status"
   Rectangle "矩形_2" at 480,205 size 60x163
      Appearance <- "Z02_Status"
   Rectangle "矩形_6" at 920,205 size 60x163
      Appearance <- "Z02_Status"
   Button "按钮_15" at 720,19 size 200x163; TextOff '工作位'
      on Press: function_b14e0dd5("Z01_Cmd", 0)
      Appearance <- "Z01_Status"
   Button "按钮_21" at 12,19 size 468x163; TextOff '******* 基本位Z1'; TextList "Cylinder_Name"
      on Press: function_b14e0dd5("Z01_Cmd", 1)
      Appearance <- "Z01_Status"
      ProcessValue <- "手动控制\CylinderIndex1"
   SymbolicIOField "符号 IO 域_9" at 546,99 size 164x83; TextOn '1'; TextOff '0'; TextList "Cylinder_QRet"
      ProcessValue <- "手动控制\CylinderIndex1"
      Appearance <- "Z01_Status"
   SymbolicIOField "符号 IO 域_10" at 986,99 size 164x83; TextOn '1'; TextOff '0'; TextList "Cylinder_QExt"
      ProcessValue <- "手动控制\CylinderIndex1"
      Appearance <- "Z01_Status"
   Rectangle "矩形_3" at 480,19 size 60x163
      Appearance <- "Z01_Status"
   Rectangle "矩形_7" at 920,19 size 60x163
      Appearance <- "Z01_Status"
   Button "按钮_16" at 720,397 size 200x163; TextOff '工作位'
      on Press: function_b14e0dd5("Z03_CmdW", 0)
      Appearance <- "Z03_Status"
   Button "按钮_23" at 12,397 size 468x163; TextOff '******* 基本位Z1'; TextList "Cylinder_Name"
      on Press: function_b14e0dd5("Z03_CmdW", 1)
      Appearance <- "Z03_Status"
      ProcessValue <- "手动控制\CylinderIndex3"
   SymbolicIOField "符号 IO 域_12" at 546,476 size 164x83; TextOn '1'; TextOff '0'; TextList "Cylinder_QRet"
      ProcessValue <- "手动控制\CylinderIndex3"
      Appearance <- "Z03_Status"
   SymbolicIOField "符号 IO 域_13" at 986,476 size 164x83; TextOn '1'; TextOff '0'; TextList "Cylinder_QExt"
      ProcessValue <- "手动控制\CylinderIndex3"
      Appearance <- "Z03_Status"
   Rectangle "矩形_4" at 480,397 size 60x163
      Appearance <- "Z03_Status"
   Rectangle "矩形_8" at 920,397 size 60x163
      Appearance <- "Z03_Status"
   Button "按钮_17" at 720,587 size 200x163; TextOff '工作位'
      on Press: function_b14e0dd5("Z04_CmdW", 0)
      Appearance <- "Z04_Status"
   Button "按钮_24" at 12,587 size 468x163; TextOff '******* 基本位Z1'; TextList "Cylinder_Name"
      on Press: function_b14e0dd5("Z04_CmdW", 1)
      Appearance <- "Z04_Status"
      ProcessValue <- "手动控制\CylinderIndex4"
   SymbolicIOField "符号 IO 域_15" at 546,667 size 164x83; TextOn '1'; TextOff '0'; TextList "Cylinder_QRet"
      ProcessValue <- "手动控制\CylinderIndex4"
      Appearance <- "Z04_Status"
   SymbolicIOField "符号 IO 域_16" at 986,667 size 164x83; TextOn '1'; TextOff '0'; TextList "Cylinder_QExt"
      ProcessValue <- "手动控制\CylinderIndex4"
      Appearance <- "Z04_Status"
   Rectangle "矩形_5" at 480,587 size 60x163
      Appearance <- "Z04_Status"
   Rectangle "矩形_9" at 920,587 size 60x163
      Appearance <- "Z04_Status"
   Button "按钮_18" at 720,777 size 200x163; TextOff '工作位'
      on Press: function_b14e0dd5("Z05_CmdW", 0)
      Appearance <- "Z05_Status"
   Button "按钮_26" at 12,777 size 468x163; TextOff '******* 基本位Z1'; TextList "Cylinder_Name"
      on Press: function_b14e0dd5("Z05_CmdW", 1)
      Appearance <- "Z05_Status"
      ProcessValue <- "手动控制\CylinderIndex5"
   SymbolicIOField "符号 IO 域_18" at 546,855 size 164x83; TextOn '1'; TextOff '0'; TextList "Cylinder_QRet"
      ProcessValue <- "手动控制\CylinderIndex5"
      Appearance <- "Z05_Status"
   SymbolicIOField "符号 IO 域_19" at 986,855 size 164x83; TextOn '1'; TextOff '0'; TextList "Cylinder_QExt"
      ProcessValue <- "手动控制\CylinderIndex5"
      Appearance <- "Z05_Status"
   Rectangle "矩形_10" at 480,777 size 60x163
      Appearance <- "Z05_Status"
   Rectangle "矩形_11" at 920,777 size 60x163
      Appearance <- "Z05_Status"
   SymbolicIOField "符号 IO 域_2" at 546,205 size 164x83; TextOn '1'; TextOff '0'; TextList "Cylinder_IRet"
      ProcessValue <- "手动控制\CylinderIndex2"
      Appearance <- "Z02_Status"
   SymbolicIOField "符号 IO 域_8" at 986,205 size 164x83; TextOn '1'; TextOff '0'; TextList "Cylinder_IExt"
      ProcessValue <- "手动控制\CylinderIndex2"
      Appearance <- "Z02_Status"
   SymbolicIOField "符号 IO 域_3" at 546,19 size 164x83; TextOn '1'; TextOff '0'; TextList "Cylinder_IRet"
      ProcessValue <- "手动控制\CylinderIndex1"
      Appearance <- "Z01_Status"
   SymbolicIOField "符号 IO 域_11" at 986,19 size 164x83; TextOn '1'; TextOff '0'; TextList "Cylinder_IExt"
      ProcessValue <- "手动控制\CylinderIndex1"
      Appearance <- "Z01_Status"
   SymbolicIOField "符号 IO 域_4" at 546,397 size 164x83; TextOn '1'; TextOff '0'; TextList "Cylinder_IRet"
      ProcessValue <- "手动控制\CylinderIndex3"
      Appearance <- "Z03_Status"
   SymbolicIOField "符号 IO 域_14" at 986,397 size 164x83; TextOn '1'; TextOff '0'; TextList "Cylinder_IExt"
      ProcessValue <- "手动控制\CylinderIndex3"
      Appearance <- "Z03_Status"
   SymbolicIOField "符号 IO 域_5" at 546,587 size 164x83; TextOn '1'; TextOff '0'; TextList "Cylinder_IRet"
      ProcessValue <- "手动控制\CylinderIndex4"
      Appearance <- "Z04_Status"
   SymbolicIOField "符号 IO 域_17" at 986,587 size 164x83; TextOn '1'; TextOff '0'; TextList "Cylinder_IExt"
      ProcessValue <- "手动控制\CylinderIndex4"
      Appearance <- "Z04_Status"
   SymbolicIOField "符号 IO 域_20" at 546,777 size 164x83; TextOn '1'; TextOff '0'; TextList "Cylinder_IRet"
      ProcessValue <- "手动控制\CylinderIndex5"
      Appearance <- "Z05_Status"
   SymbolicIOField "符号 IO 域_21" at 986,777 size 164x83; TextOn '1'; TextOff '0'; TextList "Cylinder_IExt"
      ProcessValue <- "手动控制\CylinderIndex5"
      Appearance <- "Z05_Status"

screen "198-标准通断控制_1" 1280x1024, template "Template"
   TextField "文本域_160" at 118,69 size 1040x75; Text '标准通断控制 / 伺服点动'
   SymbolicIOField "符号 IO 域_1" at 118,949 size 1040x69; TextOn '1'; TextOff '0'; TextList "操作提示"
      ProcessValue <- "DB_Message_PromptValue"
   Button "按钮_14" at 652,320 size 288x139; TextOff '工作位'
      on Press: function_b14e0dd5("Z02_CmdW", 0)
      Appearance <- "Z02_Status"
   Button "按钮_20" at 130,320 size 288x139; TextOff '******* 基本位Z1'
      on Press: function_b14e0dd5("Z02_CmdW", 1)
      Appearance <- "Z02_Status"
   SymbolicIOField "符号 IO 域_6" at 482,388 size 144x69; TextOn '1'; TextOff '0'; TextList "Cylinder_QRet"
      ProcessValue <- "手动控制\CylinderIndex2"
      Appearance <- "Z02_Status"
   SymbolicIOField "符号 IO 域_7" at 1002,388 size 148x69; TextOn '1'; TextOff '0'; TextList "Cylinder_QExt"
      ProcessValue <- "手动控制\CylinderIndex2"
      Appearance <- "Z02_Status"
   Rectangle "矩形_2" at 422,323 size 54x132
      Appearance <- "Z02_Status"
   Rectangle "矩形_6" at 944,323 size 54x132
      Appearance <- "Z02_Status"
   Button "按钮_15" at 652,163 size 288x137; TextOff '工作位'
      on Press: function_b14e0dd5("Z01_Cmd", 0)
      Appearance <- "Z01_Status"
   Button "按钮_21" at 130,163 size 288x137; TextOff '******* 基本位Z1'
      on Press: function_b14e0dd5("Z01_Cmd", 1)
      Appearance <- "Z01_Status"
   SymbolicIOField "符号 IO 域_9" at 482,228 size 144x69; TextOn '1'; TextOff '0'; TextList "Cylinder_QRet"
      ProcessValue <- "手动控制\CylinderIndex1"
      Appearance <- "Z01_Status"
   SymbolicIOField "符号 IO 域_10" at 1002,228 size 148x69; TextOn '1'; TextOff '0'; TextList "Cylinder_QExt"
      ProcessValue <- "手动控制\CylinderIndex1"
      Appearance <- "Z01_Status"
   Rectangle "矩形_3" at 422,163 size 54x132
      Appearance <- "Z01_Status"
   Rectangle "矩形_7" at 944,163 size 54x132
      Appearance <- "Z01_Status"
   SymbolicIOField "符号 IO 域_2" at 482,320 size 144x69; TextOn '1'; TextOff '0'; TextList "Cylinder_IRet"
      ProcessValue <- "手动控制\CylinderIndex2"
      Appearance <- "Z02_Status"
   SymbolicIOField "符号 IO 域_8" at 1002,320 size 148x69; TextOn '1'; TextOff '0'; TextList "Cylinder_IExt"
      ProcessValue <- "手动控制\CylinderIndex2"
      Appearance <- "Z02_Status"
   SymbolicIOField "符号 IO 域_3" at 482,163 size 144x69; TextOn '1'; TextOff '0'; TextList "Cylinder_IRet"
      ProcessValue <- "手动控制\CylinderIndex1"
      Appearance <- "Z01_Status"
   SymbolicIOField "符号 IO 域_11" at 1002,163 size 148x69; TextOn '1'; TextOff '0'; TextList "Cylinder_IExt"
      ProcessValue <- "手动控制\CylinderIndex1"
      Appearance <- "Z01_Status"
   Button "按钮_1" at 652,476 size 288x139; TextOff '工作位'
      on Press: function_b14e0dd5("Z02_CmdW", 0)
      Appearance <- "Z02_Status"
   Button "按钮_2" at 130,476 size 288x139; TextOff '******* 基本位Z1'
      on Press: function_b14e0dd5("Z02_CmdW", 1)
      Appearance <- "Z02_Status"
   SymbolicIOField "符号 IO 域_4" at 482,544 size 144x69; TextOn '1'; TextOff '0'; TextList "Cylinder_QRet"
      ProcessValue <- "手动控制\CylinderIndex2"
      Appearance <- "Z02_Status"
   SymbolicIOField "符号 IO 域_5" at 1002,544 size 148x69; TextOn '1'; TextOff '0'; TextList "Cylinder_QExt"
      ProcessValue <- "手动控制\CylinderIndex2"
      Appearance <- "Z02_Status"
   Rectangle "矩形" at 422,477 size 54x132
      Appearance <- "Z02_Status"
   Rectangle "矩形_4" at 944,477 size 54x132
      Appearance <- "Z02_Status"
   SymbolicIOField "符号 IO 域_12" at 482,476 size 144x69; TextOn '1'; TextOff '0'; TextList "Cylinder_IRet"
      ProcessValue <- "手动控制\CylinderIndex2"
      Appearance <- "Z02_Status"
   SymbolicIOField "符号 IO 域_13" at 1002,476 size 148x69; TextOn '1'; TextOff '0'; TextList "Cylinder_IExt"
      ProcessValue <- "手动控制\CylinderIndex2"
      Appearance <- "Z02_Status"

screen "199-标准通断模板_2" 1280x1024, template "Template"
   TextField "文本域_160" at 118,69 size 1040x75; Text '标准通断控制 / 伺服点动'
   SymbolicIOField "符号 IO 域_1" at 118,949 size 1040x69; TextOn '1'; TextOff '0'; TextList "操作提示"
      ProcessValue <- "DB_Message_PromptValue"
   Group "Group" at 130,163 size 1020x777
   Button "按钮_14" at 652,320 size 288x139; TextOff '工作位'
      on Press: function_b14e0dd5("Z02_CmdW", 0)
      Appearance <- "Z02_Status"
   Button "按钮_20" at 130,320 size 288x139; TextOff '******* 基本位Z1'
      on Press: function_b14e0dd5("Z02_CmdW", 1)
      Appearance <- "Z02_Status"
   SymbolicIOField "符号 IO 域_6" at 482,388 size 144x69; TextOn '1'; TextOff '0'; TextList "Cylinder_QRet"
      ProcessValue <- "手动控制\CylinderIndex2"
      Appearance <- "Z02_Status"
   SymbolicIOField "符号 IO 域_7" at 1002,388 size 148x69; TextOn '1'; TextOff '0'; TextList "Cylinder_QExt"
      ProcessValue <- "手动控制\CylinderIndex2"
      Appearance <- "Z02_Status"
   Rectangle "矩形_2" at 422,323 size 54x132
      Appearance <- "Z02_Status"
   Rectangle "矩形_6" at 944,323 size 54x132
      Appearance <- "Z02_Status"
   Button "按钮_15" at 652,163 size 288x137; TextOff '工作位'
      on Press: function_b14e0dd5("Z01_Cmd", 0)
      Appearance <- "Z01_Status"
   Button "按钮_21" at 130,163 size 288x137; TextOff '******* 基本位Z1'
      on Press: function_b14e0dd5("Z01_Cmd", 1)
      Appearance <- "Z01_Status"
   SymbolicIOField "符号 IO 域_9" at 482,228 size 144x69; TextOn '1'; TextOff '0'; TextList "Cylinder_QRet"
      ProcessValue <- "手动控制\CylinderIndex1"
      Appearance <- "Z01_Status"
   SymbolicIOField "符号 IO 域_10" at 1002,228 size 148x69; TextOn '1'; TextOff '0'; TextList "Cylinder_QExt"
      ProcessValue <- "手动控制\CylinderIndex1"
      Appearance <- "Z01_Status"
   Rectangle "矩形_3" at 422,163 size 54x132
      Appearance <- "Z01_Status"
   Rectangle "矩形_7" at 944,163 size 54x132
      Appearance <- "Z01_Status"
   Button "按钮_16" at 652,480 size 288x139; TextOff '工作位'
      on Press: function_b14e0dd5("Z03_CmdW", 0)
      Appearance <- "Z03_Status"
   Button "按钮_23" at 130,480 size 288x139; TextOff '******* 基本位Z1'
      on Press: function_b14e0dd5("Z03_CmdW", 1)
      Appearance <- "Z03_Status"
   SymbolicIOField "符号 IO 域_12" at 482,548 size 144x69; TextOn '1'; TextOff '0'; TextList "Cylinder_QRet"
      ProcessValue <- "手动控制\CylinderIndex3"
      Appearance <- "Z03_Status"
   SymbolicIOField "符号 IO 域_13" at 1002,548 size 148x69; TextOn '1'; TextOff '0'; TextList "Cylinder_QExt"
      ProcessValue <- "手动控制\CylinderIndex3"
      Appearance <- "Z03_Status"
   Rectangle "矩形_4" at 422,483 size 54x132
      Appearance <- "Z03_Status"
   Rectangle "矩形_8" at 944,483 size 54x132
      Appearance <- "Z03_Status"
   Button "按钮_17" at 652,643 size 288x137; TextOff '工作位'
      on Press: function_b14e0dd5("Z04_CmdW", 0)
      Appearance <- "Z04_Status"
   Button "按钮_24" at 130,643 size 288x137; TextOff '******* 基本位Z1'
      on Press: function_b14e0dd5("Z04_CmdW", 1)
      Appearance <- "Z04_Status"
   SymbolicIOField "符号 IO 域_15" at 482,708 size 144x69; TextOn '1'; TextOff '0'; TextList "Cylinder_QRet"
      ProcessValue <- "手动控制\CylinderIndex4"
      Appearance <- "Z04_Status"
   SymbolicIOField "符号 IO 域_16" at 1002,708 size 148x69; TextOn '1'; TextOff '0'; TextList "Cylinder_QExt"
      ProcessValue <- "手动控制\CylinderIndex4"
      Appearance <- "Z04_Status"
   Rectangle "矩形_5" at 422,643 size 54x132
      Appearance <- "Z04_Status"
   Rectangle "矩形_9" at 944,643 size 54x132
      Appearance <- "Z04_Status"
   Button "按钮_18" at 652,803 size 288x137; TextOff '工作位'
      on Press: function_b14e0dd5("Z05_CmdW", 0)
      Appearance <- "Z05_Status"
   Button "按钮_26" at 130,803 size 288x137; TextOff '******* 基本位Z1'
      on Press: function_b14e0dd5("Z05_CmdW", 1)
      Appearance <- "Z05_Status"
   SymbolicIOField "符号 IO 域_18" at 482,868 size 144x69; TextOn '1'; TextOff '0'; TextList "Cylinder_QRet"
      ProcessValue <- "手动控制\CylinderIndex5"
      Appearance <- "Z05_Status"
   SymbolicIOField "符号 IO 域_19" at 1002,868 size 148x69; TextOn '1'; TextOff '0'; TextList "Cylinder_QExt"
      ProcessValue <- "手动控制\CylinderIndex5"
      Appearance <- "Z05_Status"
   Rectangle "矩形_10" at 422,803 size 54x131
      Appearance <- "Z05_Status"
   Rectangle "矩形_11" at 944,804 size 54x131
      Appearance <- "Z05_Status"
   SymbolicIOField "符号 IO 域_2" at 482,320 size 144x69; TextOn '1'; TextOff '0'; TextList "Cylinder_IRet"
      ProcessValue <- "手动控制\CylinderIndex2"
      Appearance <- "Z02_Status"
   SymbolicIOField "符号 IO 域_8" at 1002,320 size 148x69; TextOn '1'; TextOff '0'; TextList "Cylinder_IExt"
      ProcessValue <- "手动控制\CylinderIndex2"
      Appearance <- "Z02_Status"
   SymbolicIOField "符号 IO 域_3" at 482,163 size 144x69; TextOn '1'; TextOff '0'; TextList "Cylinder_IRet"
      ProcessValue <- "手动控制\CylinderIndex1"
      Appearance <- "Z01_Status"
   SymbolicIOField "符号 IO 域_11" at 1002,163 size 148x69; TextOn '1'; TextOff '0'; TextList "Cylinder_IExt"
      ProcessValue <- "手动控制\CylinderIndex1"
      Appearance <- "Z01_Status"
   SymbolicIOField "符号 IO 域_4" at 482,480 size 144x69; TextOn '1'; TextOff '0'; TextList "Cylinder_IRet"
      ProcessValue <- "手动控制\CylinderIndex3"
      Appearance <- "Z03_Status"
   SymbolicIOField "符号 IO 域_14" at 1002,480 size 148x69; TextOn '1'; TextOff '0'; TextList "Cylinder_IExt"
      ProcessValue <- "手动控制\CylinderIndex3"
      Appearance <- "Z03_Status"
   SymbolicIOField "符号 IO 域_5" at 482,643 size 144x69; TextOn '1'; TextOff '0'; TextList "Cylinder_IRet"
      ProcessValue <- "手动控制\CylinderIndex4"
      Appearance <- "Z04_Status"
   SymbolicIOField "符号 IO 域_17" at 1002,643 size 148x69; TextOn '1'; TextOff '0'; TextList "Cylinder_IExt"
      ProcessValue <- "手动控制\CylinderIndex4"
      Appearance <- "Z04_Status"
   SymbolicIOField "符号 IO 域_20" at 482,803 size 144x69; TextOn '1'; TextOff '0'; TextList "Cylinder_IRet"
      ProcessValue <- "手动控制\CylinderIndex5"
      Appearance <- "Z05_Status"
   SymbolicIOField "符号 IO 域_21" at 1002,803 size 148x69; TextOn '1'; TextOff '0'; TextList "Cylinder_IExt"
      ProcessValue <- "手动控制\CylinderIndex5"
      Appearance <- "Z05_Status"

Template "Template" 1280x1024
   Button "Template_模板_按钮_22" at 1158,829 size 120x192; TextOn '运行 设置'; TextOff '报警 信息'
      on Release: function_dbe01993("DB_SysMode_TPSetPageNo", 1, "DB_SysMode_TPCurPageType", "DB_SysMode_TPCurSubPage"); ActivateScreenByNumber("DB_SysMode_TPSetPageNo", 0)
      on Press: SetTag("DB_SysMode_TPCurPageType", 9); SetTag("DB_SysMode_TPCurSubPage", 0)
      Appearance <- "DB_SysMode_TPCurPageType"
   Button "Template_模板_按钮_23" at 1158,68 size 120x192; TextOn '运行 设置'; TextOff '手动 画面'
      on Release: function_dbe01993("DB_SysMode_TPSetPageNo", 1, "DB_SysMode_TPCurPageType", "DB_SysMode_TPCurSubPage"); ActivateScreenByNumber("DB_SysMode_TPSetPageNo", 0)
      on Press: SetTag("DB_SysMode_TPCurPageType", 100); SetTag("DB_SysMode_TPCurSubPage", 0)
      Appearance <- "DB_SysMode_TPCurPageType"
   Button "Template_模板_按钮_24" at 1158,260 size 120x192; TextOn '运行 设置'; TextOff '自动 监视'
      on Activate: function_bed61462(2)
      on Release: function_dbe01993("DB_SysMode_TPSetPageNo", 1, "DB_SysMode_TPCurPageType", "DB_SysMode_TPCurSubPage"); ActivateScreenByNumber("DB_SysMode_TPSetPageNo", 0)
      on Press: SetTag("DB_SysMode_TPCurPageType", 200); SetTag("DB_SysMode_TPCurSubPage", 0)
      Appearance <- "DB_SysMode_TPCurPageType"
   Button "Template_模板_按钮_25" at 1158,452 size 120x192; TextOn '运行 设置'; TextOff '参数 设置'; Authorization "Operate"
      on Release: function_dbe01993("DB_SysMode_TPSetPageNo", 1, "DB_SysMode_TPCurPageType", "DB_SysMode_TPCurSubPage"); ActivateScreenByNumber("DB_SysMode_TPSetPageNo", 0)
      on Press: SetTag("DB_SysMode_TPCurPageType", 300); SetTag("DB_SysMode_TPCurSubPage", 0); function_b3f726e6("DB_Parameter_TP_Cmd", 2)
      Appearance <- "DB_SysMode_TPCurPageType"
   Button "Template_模板_按钮_19" at 1158,644 size 120x192; TextOn '运行 设置'; TextOff '型号 选择'
      on Release: function_dbe01993("DB_SysMode_TPSetPageNo", 1, "DB_SysMode_TPCurPageType", "DB_SysMode_TPCurSubPage"); ActivateScreenByNumber("DB_SysMode_TPSetPageNo", 0)
      on Press: SetTag("DB_SysMode_TPCurPageType", 400); SetTag("DB_SysMode_TPCurSubPage", 0)
      Appearance <- "DB_SysMode_TPSetPageNo"
   Button "Template_模板_按钮_32" at 0,68 size 120x192; TextOn '运行 设置'; TextOff '手动 画面'; TextList "按钮1"
      on Release: function_dbe01993("DB_SysMode_TPSetPageNo", 1, "DB_SysMode_TPCurPageType", "DB_SysMode_TPCurSubPage"); ActivateScreenByNumber("DB_SysMode_TPSetPageNo", 0)
      on Press: SetTag("DB_SysMode_TPCurSubPage", 0)
      Appearance <- "DB_SysMode_TPCurSubPage"
      ProcessValue <- "DB_SysMode_TPCurPageType"
   Button "Template_模板_按钮_35" at 0,260 size 120x192; TextOn '运行 设置'; TextOff '手动 画面'; TextList "按钮2"
      on Release: function_dbe01993("DB_SysMode_TPSetPageNo", 1, "DB_SysMode_TPCurPageType", "DB_SysMode_TPCurSubPage"); ActivateScreenByNumber("DB_SysMode_TPSetPageNo", 0)
      on Press: SetTag("DB_SysMode_TPCurSubPage", 20)
      Appearance <- "DB_SysMode_TPCurSubPage"
      ProcessValue <- "DB_SysMode_TPCurPageType"
   Button "Template_模板_按钮_36" at 0,452 size 120x192; TextOn '运行 设置'; TextOff '手动 画面'; TextList "按钮3"
      on Release: function_dbe01993("DB_SysMode_TPSetPageNo", 1, "DB_SysMode_TPCurPageType", "DB_SysMode_TPCurSubPage"); ActivateScreenByNumber("DB_SysMode_TPSetPageNo", 0)
      on Press: SetTag("DB_SysMode_TPCurSubPage", 40)
      Appearance <- "DB_SysMode_TPCurSubPage"
      ProcessValue <- "DB_SysMode_TPCurPageType"
   Button "Template_模板_按钮_37" at 0,832 size 120x192; TextOn '运行 设置'; TextOff '手动 画面'; TextList "按钮4"
      on Release: function_dbe01993("DB_SysMode_TPSetPageNo", 1, "DB_SysMode_TPCurPageType", "DB_SysMode_TPCurSubPage"); ActivateScreenByNumber("DB_SysMode_TPSetPageNo", 0)
      on Press: SetTag("DB_SysMode_TPCurSubPage", 60)
      Appearance <- "DB_SysMode_TPCurSubPage"
      ProcessValue <- "DB_SysMode_TPCurPageType"
   DateTimeField "模板_日期/时间域_1" at 594,0 size 683x69
      ProcessValue <- "DB_SysMode_Sys_Time_CurPLCTime"
   Button "Template_模板_按钮_3" at 1126,1 size 149x66; TextOn '运行 设置'; TextOff '最小化 手动 画面'; TextList "按钮1"
      on Press: function_bed61462(4)
      ProcessValue <- "DB_SysMode_TPCurPageType"
   Button "Template_模板_按钮_4" at 975,1 size 149x66; TextOn '运行 设置'; TextOff '退出 手动 画面'; TextList "按钮1"
      on Press: StopRuntime(0)
      ProcessValue <- "DB_SysMode_TPCurPageType"
   Button "Template_模板_按钮_1" at 0,645 size 120x192; TextOff '气缸 操作'
      on Release: ActivateScreen("190-气缸控制", 0)
      on Press: SetTag("DB_SysMode_TPSetPageNo", 190); SetTag("Cylinder_Index_Max", 12); SetTag("Cylinder_Index_Min", 1); SetTag("DB_SysMode_Cylinder_Index", 1)
      Appearance <- "DB_SysMode_TPCurSubPage"
   TextField "文本域_1" at 0,0 size 594x69; Text '电锤 功能测试 / TMAP——ManualOperation'

screen "100-KUKA机器人手动操作" 1280x1024, template "Template"
   Button "按钮_4" at 130,550 size 145x77; TextOff 'CCD Trige / 批头校验'; Authorization "User administration"
      on Press: function_b14e0dd5("DB_KuKa_MainCtrl.CheckAiguille.StartCmd", 0)
      Appearance <- "DB_KuKa_MainCtrl.CheckAiguille.StepStart"
   Button "按钮_5" at 777,550 size 145x77; TextOff 'CCD Trige / 水平钻孔'; Authorization "User administration"
      on Press: function_b14e0dd5("DB_KuKa_MainCtrl.DrillHorizontal.StartCmd", 0)
      Appearance <- "DB_KuKa_MainCtrl.DrillHorizontal.StepStart"
   Button "按钮_12" at 281,648 size 145x77; TextOff 'CCD Trige / 清洁'; Authorization "User administration"
      on Press: function_b14e0dd5("DB_KuKa_MainCtrl.CleanTool.StartCmd", 0)
      Appearance <- "DB_KuKa_MainCtrl.CleanTool.StepStart"
   SymbolicIOField "符号 IO 域_2" at 122,951 size 1040x64; TextOn '1'; TextOff '0'; TextList "操作提示"
      ProcessValue <- "DB_Message_PromptValue"
   Group "Group" at 126,153 size 1021x320; Authorization "User administration"
   Button "按钮_6" at 130,648 size 145x77; TextOff 'CCD Trige / 换夹具'; Authorization "User administration"
      on Press: function_b14e0dd5("DB_KuKa_MainCtrl.ChangeTool.StartCmd", 0)
      Appearance <- "DB_KuKa_MainCtrl.ChangeTool.StepStart"
   Button "按钮_8" at 469,550 size 145x77; TextOff 'CCD Trige / 向下钻孔'; Authorization "User administration"
      on Press: function_b14e0dd5("DB_KuKa_MainCtrl.DrillDownload.StartCmd", 0)
      Appearance <- "DB_KuKa_MainCtrl.DrillDownload.StepStart"
   Button "按钮_9" at 624,550 size 145x77; TextOff 'CCD Trige / 向上钻孔'; Authorization "User administration"
      on Press: function_b14e0dd5("DB_KuKa_MainCtrl.DrillUpload.StartCmd", 0)
      Appearance <- "DB_KuKa_MainCtrl.DrillUpload.StepStart"
   IOField "I/O field_5" at 565,858 size 141x47; FormatPattern 99.9999
      ProcessValue <- "DB_Component_Aux_Pressure"
   TextField "文本域" at 713,857 size 65x48; Text 'MPa'
   SymbolicIOField "符号 I/O 域_1" at 280,552 size 146x66; TextOff '0'; TextOn '1'; TextList "校验"
      ProcessValue <- "DB_KuKa_MainCtrl.Aux.CheckNo"
   IOField "I/O field_6" at 565,807 size 141x47; FormatPattern 9999.99
      ProcessValue <- "DB_Timer_Force"
   TextField "文本域_1" at 713,806 size 65x48; Text 'N'
   Button "按钮_14" at 998,809 size 147x113; TextOff 'ST02伺服 点动前进 返回'; TextList "Cylinder_Name_1"
      on Press: function_efd93a16()
      ProcessValue <- "CylinderIndex1"
   TextField "Text field_10" at 679,215 size 175x64; Text 'JobNO / 选择动作'
   TextField "Text field_1" at 251,406 size 120x67; Text 'TaskDone / 完成'
      Appearance <- "DB_Component_Robot_TP_Status"
   TextField "Text field_3" at 377,406 size 120x67; Text 'TaskIO / 合格'
      Appearance <- "DB_Component_Robot_TP_Status"
   TextField "Text field_4" at 503,406 size 120x67; Text 'TaskNIO / 失败'
      Appearance <- "DB_Component_Robot_TP_Status"
   TextField "Text field_5" at 628,406 size 120x67; Text 'JobOK / 原点'
      Appearance <- "DB_Component_Robot_TP_Status"
   TextField "Text field_7" at 126,406 size 120x67; Text 'Busy / 运行'
      Appearance <- "DB_Component_Robot_TP_Status"
   Button "按钮_2" at 127,215 size 179x130; TextOff 'CCD Trige / 启动'; Authorization "User administration"
   SymbolicIOField "符号 IO 域_1" at 126,345 size 1021x58; TextOn '1'; TextOff '0'; TextList "KuKaRobotStatusPrompt"
      ProcessValue <- "DB_Component_Robot_Status_PromptValue"
      Appearance <- "DB_Component_Robot_Status_PromptValue"
   TextField "Text field_2" at 754,406 size 120x67; Text 'Ready'
      Appearance <- "DB_Component_Robot_TP_Status"
   TextField "Text field_8" at 880,406 size 120x67; Text 'xx'
   TextField "文本域_5" at 127,153 size 997x59; Text '伺服点动 / KUKA机器人'
   IOField "I/O field_2" at 1006,282 size 141x61; FormatPattern 999
      ProcessValue <- "DB_Component_Robot_CTRL_OUT_ProgNo"
   TextField "Text field_9" at 1006,215 size 141x64; Text 'JobNO / 反馈程序号'
   IOField "I/O field_4" at 1030,156 size 117x49; FormatPattern 99999
      ProcessValue <- "DB_Component_Robot_Step_Main"
      Visibility <- "DB_Component_Robot_Step_Main"
   Button "按钮_1" at 311,215 size 179x130; TextOff 'CCD Trige / 回原点'
      on Press: function_b14e0dd5("DB_Component_Robot_TP_Cmd", 9)
   Button "按钮_3" at 495,215 size 179x130; TextOff 'CCD Trige / 停止'
      on Press: function_b14e0dd5("DB_Component_Robot_TP_Cmd", 10)
   IOField "IO 域_11" at 1006,406 size 141x67; FormatPattern 999999; Unit s
      ProcessValue <- "DB_Component_Robot_CTRL_OUT_LastCylceTime"
   SymbolicIOField "Symbolic I/O field_2" at 679,282 size 175x61; TextOn '111'; TextOff '1111'; TextList "机器人动作号"
      ProcessValue <- "AG1520RobotIndex"
   IOField "I/O field_1" at 859,282 size 141x61; FormatPattern 999
      ProcessValue <- "DB_Component_Robot_CTRL_IN_ProgNo"
   TextField "Text field_6" at 859,215 size 141x64; Text 'JobNO / 输入程序号'
   IOField "I/O field_3" at 127,156 size 117x49; FormatPattern 99999
      ProcessValue <- "DB_Component_Robot_CTRL_OUT_ErrorCode"
      Appearance <- "DB_Component_Robot_CTRL_OUT_ErrorCode"
   Button "按钮_7" at 141,811 size 170x90; TextOff '位移传感器 标定界面'
      on Press: SetTag("DB_AddrRegister_Analog_IN_V4_FBCall_IndexNO", 1); SetTag("DB_AddrRegister_Analog_IN_V4_FBCall_StartAddr", 722); SetTag("ObjectComment", '移传感器标定界面'); SetTag("Object_Description", '模拟量输入信号：IW88,单位mm'); ActivateScreen("385-模拟量输入_V4", 0)
   Button "按钮_10" at 360,811 size 170x90; TextOff '模拟量 输出标定'
      on Press: SetTag("Object_Description", '伺服比例阀模拟量输出信号：QW88,单位bar;'); ActivateScreen("386-模拟量输出_V3", 0)
   Button "按钮_11" at 807,811 size 170x90; TextOff '气缸压力 标定界面'
      on Press: SetTag("DB_AddrRegister_Analog_IN_V4_FBCall_IndexNO", 1); SetTag("DB_AddrRegister_Analog_IN_V4_FBCall_StartAddr", 522); SetTag("ObjectComment", '气缸压力标定界面'); SetTag("Object_Description", '模拟量输入信号：IW88,单位mm'); ActivateScreen("385-模拟量输入_V4", 0)

screen "385-模拟量输入_V4" 1280x1024, template "Template"
   Button "按钮_8" at 653,811 size 248x122; TextOff '保 存'
      on Press: function_b14e0dd5("DB_Parameter_TP_Cmd", 8)
      Appearance <- "DB_Parameter_TP_Status"
   Button "按钮_3" at 907,811 size 243x122; TextOff '返 回'
      on Press: function_efd93a16()
   Group "Group" at 123,103 size 1026x544
   SymbolicIOField "符号 IO 域_1" at 123,951 size 1040x64; TextOn '1'; TextOff '0'; TextList "操作提示"
      ProcessValue <- "DB_Message_PromptValue"
   IOField "I/O field_5" at 123,103 size 1026x58; FormatPattern ????????????????????????????????????????????????????????????????????????????????
      ProcessValue <- "ObjectComment"
   Button "按钮_6" at 846,327 size 300x76; TextOff '根据PreSet计算偏置'
      on Press: function_b14e0dd5("Analog_In_V4_TP_Cmd", 8)
      Appearance <- "Analog_In_V4_TP_Cmd"
   TextField "Text field_2" at 126,327 size 132x76; Text 'Gain:'
   IOField "I/O field_6" at 262,327 size 105x76
      ProcessValue <- "Analog_In_V4_Ctrl_IN_TP_AI_Gain"
   TextField "Text field_4" at 849,171 size 159x74; Text 'CurValue:'
   IOField "I/O field_7" at 1013,171 size 132x74; FormatPattern 9999.999
      ProcessValue <- "Analog_In_V4_Ctrl_Out_Cur_Val_Out"
   TextField "Text field_7" at 373,327 size 126x76; Text 'OffSet'
   IOField "I/O field_8" at 501,327 size 107x76
      ProcessValue <- "Analog_In_V4_Ctrl_IN_TP_AI_OffSet"
   TextField "Text field_8" at 612,327 size 119x76; Text 'PreSet:'
   IOField "I/O field_13" at 733,327 size 105x76
      ProcessValue <- "Analog_In_V4_Ctrl_IN_TP_PreSetValue"
   TextField "Text field_13" at 126,570 size 159x76; Text 'Point2:'
   IOField "I/O field_14" at 289,570 size 153x76
      ProcessValue <- "Analog_In_V4_Ctrl_IN_TP_ActualAI_2"
   TextField "Text field_14" at 126,488 size 159x76; Text 'Point1:'
   IOField "I/O field_15" at 289,488 size 153x76
      ProcessValue <- "Analog_In_V4_Ctrl_IN_TP_ActualAI_1"
   TextField "Text field_15" at 681,570 size 159x76; Text 'Actual:'
   IOField "I/O field_16" at 846,570 size 153x76; FormatPattern 99999.999
      ProcessValue <- "Analog_In_V4_Ctrl_IN_TP_ActualAI_Value2"
   TextField "Text field_16" at 681,488 size 159x76; Text 'Actual:'
   IOField "I/O field_17" at 846,488 size 153x76; FormatPattern 99999.999
      ProcessValue <- "Analog_In_V4_Ctrl_IN_TP_ActualAI_Value1"
   Button "按钮_7" at 1007,488 size 139x159; TextOff '计算 增益及偏置'
      on Press: function_b14e0dd5("Analog_In_V4_TP_Cmd", 11)
      Appearance <- "Analog_In_V4_TP_Cmd"
   Button "按钮_9" at 448,488 size 226x78; TextOff 'ReadPLCValue'
      on Press: function_b14e0dd5("Analog_In_V4_TP_Cmd", 9)
      Appearance <- "Analog_In_V4_TP_Cmd"
   Button "按钮_10" at 448,568 size 226x78; TextOff 'ReadPLCValue'
      on Press: function_b14e0dd5("Analog_In_V4_TP_Cmd", 10)
      Appearance <- "Analog_In_V4_TP_Cmd"
   TextField "文本域_7" at 126,411 size 1019x74; Text '标定方法2，两点标定'
   TextField "文本域_8" at 126,250 size 1019x74; Text '标定方法1，根据量程Gain及PreSet计算偏置OffSet, 计算公式： y=Gain*AI+ OffSet'
   IOField "I/O field_1" at 126,173 size 716x71; FormatPattern ????????????????????????????????????????????????????????????????????????????????
      ProcessValue <- "Object_Description"

screen "386-模拟量输出_V3" 1280x1024, template "Template"
   Button "按钮_8" at 653,811 size 248x122; TextOff '保 存'
      on Press: function_b14e0dd5("DB_Parameter_TP_Cmd", 8)
      Appearance <- "DB_Parameter_TP_Status"
   Button "按钮_3" at 907,811 size 243x122; TextOff '返 回'
      on Press: function_efd93a16()
   SymbolicIOField "符号 IO 域_1" at 123,951 size 1040x64; TextOn '1'; TextOff '0'; TextList "操作提示"
      ProcessValue <- "DB_Message_PromptValue"
   TextField "Text field_7" at 767,317 size 158x73; Text 'SetTarget:'
   IOField "I/O field_11" at 930,317 size 131x73
      ProcessValue <- "DB_Component_Analog_Out_Ctrl_IN_Target"
   TextField "Text field_13" at 134,550 size 158x75; Text 'Point2:'
   IOField "I/O field_14" at 296,550 size 166x75; FormatPattern 99999.99
      ProcessValue <- "Analog_Out_Ctrl_IN_TP_ActualAO_2"
   TextField "Text field_14" at 134,469 size 158x75; Text 'Point1:'
   IOField "I/O field_15" at 296,469 size 166x75; FormatPattern 99999.99
      ProcessValue <- "Analog_Out_Ctrl_IN_TP_ActualAO_1"
   TextField "Text field_15" at 698,550 size 158x75; Text 'Actual:'
   IOField "I/O field_16" at 861,550 size 152x75
      ProcessValue <- "Analog_Out_Ctrl_IN_TP_ActualAO_Value2"
   TextField "Text field_16" at 698,469 size 158x75; Text 'Actual:'
   IOField "I/O field_17" at 861,469 size 152x75
      ProcessValue <- "Analog_Out_Ctrl_IN_TP_ActualAO_Value1"
   Button "按钮_9" at 466,469 size 224x77; TextOff 'ReadPLCValue'
      on Press: function_b14e0dd5("DB_Component.Analog_Out_1.Cmd.Read1", 0)
      Appearance <- "DB_Component.Analog_Out_1.Cmd.Read1"
   Button "按钮_10" at 466,548 size 224x77; TextOff 'ReadPLCValue'
      on Press: function_b14e0dd5("DB_Component.Analog_Out_1.Cmd.Read2", 0)
      Appearance <- "DB_Component.Analog_Out_1.Cmd.Read2"
   TextField "文本域_3" at 134,393 size 928x73; Text '标定方法2，两点标定'
   Button "按钮_7" at 1017,468 size 139x159; TextOff '计算 增益及偏置'
      on Press: function_b14e0dd5("DB_Component.Analog_Out_1.Confirm", 0)
      Appearance <- "DB_Component.Analog_Out_1.Confirm"

VB script "LanguageChange"
   '注意：要启动脚本，请按下 <Ctrl><空格>，然后就可以看到各种不同函数。
   '通过使用系统函数或 WinCC flexible 对象模型来编写脚本。您可以通过 HMI 运行系统对象很容易地访问系统
   '。挑选对象引用的一个很便利的
   '方式是按下 <Alt><右箭头>。通过使用编程语言 VBScript 的基本功能部件
   '来设计复杂的脚本，并可以直接通过名称，例如 tag = 5，来访问变量。
   If SmartTags("Language") >=2 Then
   	SmartTags("Language")= 0
   End If

VB script "Script_2"
   '注意：要启动脚本，请按下 <Ctrl><空格>，然后就可以看到各种不同函数。'通过使用系统函数或 WinCC flexible 对象模型来编写脚本。您可以通过 HMI 运行系统对象很容易地访问系统'。挑选对象引用的一个很便利的'方式是按下 <Alt><右箭头>。通过使用编程语言 VBScript 的基本功能部件'来设计复杂的脚本，并可以直接通过名称，例如 tag = 5，来访问变量。
*)